(* IEC 61131-3 sources: daoli-st-library/DL_Process (part 16) *)

(* ---- FC_DL_RegisterErrorCalc.st ---- *)
(*
  DL Factory R83 | FC_DL_RegisterErrorCalc
  功能：把纵向与横向套准误差合成偏差幅值与方位角，并按合成允差判定超差。
  开源溯源：无（clean-room 自研，依据公开工艺公式，来源=行业通用公式，许可证=MIT，借鉴点=公式结构）
  规则：R1-R21 全遵守
*)
FUNCTION FC_DL_RegisterErrorCalc : REAL
VAR_INPUT
    fErrMd    : REAL; // 纵向（走料方向）套准误差，正=超前 [mm] / Machine-direction error [mm]
    fErrCd    : REAL; // 横向（幅宽方向）套准误差，正=右偏 [mm] / Cross-direction error [mm]
    fTolMm    : REAL; // 套准允差（合成偏差上限）[mm] / Tolerance on composite error [mm]
    fSpeedMpm : REAL; // 料带走料速度 [m/min] / Web speed [m/min]
END_VAR
VAR_OUTPUT
    fErrComp  : REAL; // 合成偏差幅值 [mm] / Composite error magnitude [mm]
    fErrAngle : REAL; // 误差方位角，0=纵向 90=横向 [°] / Error azimuth [deg]
    xOutTol   : BOOL; // 超差标志（TRUE=超差需调整）/ Out-of-tolerance flag
END_VAR
VAR
    fSq  : REAL; // 误差平方和 [mm²] / Sum of squared errors [mm^2]
    fRad : REAL; // 方位角弧度 [rad] / Azimuth in radians [rad]
    fPi  : REAL := 3.14159265358979; // 圆周率常量，弧度转度用（R19 已引用）/ Pi constant, referenced
END_VAR
// 出口预置：三出口统一预置（R256）
fErrComp := 0.0; fErrAngle := 0.0; xOutTol := FALSE;
// 非有限拦截 + 量纲自检：允差必须为正（R20/R21）
IF NOT (fErrMd > -1.0E30 AND fErrMd < 1.0E30) OR NOT (fErrCd > -1.0E30 AND fErrCd < 1.0E30) OR NOT (fTolMm > -1.0E30 AND fTolMm < 1.0E30) OR NOT (fSpeedMpm > -1.0E30 AND fSpeedMpm < 1.0E30) OR fTolMm <= 0.0 THEN
    FC_DL_RegisterErrorCalc := -1.0; RETURN;   // 哨兵 -1：非有限或允差非正 / Sentinel -1
END_IF
// 合成偏差：欧氏范数，开方前非负闸（R4）
fSq := fErrMd * fErrMd + fErrCd * fErrCd;  // 平方和 [mm²] / Sum of squares [mm^2]
IF fSq >= 0.0 THEN                  // 开方前非负闸 / Gate before square root
    fErrComp := SQRT(fSq);          // 合成偏差 [mm] / Composite error [mm]
ELSE
    fErrComp := 0.0;                // 浮点异常防御缺省 / Float anomaly default
END_IF
// 方位角：纵向分量为分母，显式零闸后取反正切，纯横向走 ±90° 分支
IF ABS(fErrMd) > 1.0E-6 THEN        // 分母零闸（R4/R21）/ Denominator zero gate
    fRad      := ATAN(fErrCd / fErrMd);   // 象限角 [-π/2, π/2] / Quadrant angle [rad]
    fErrAngle := fRad * 180.0 / fPi;      // 转度 [°] / Convert to degrees [deg]
ELSIF fErrCd >= 0.0 THEN
    fErrAngle := 90.0;              // 纯横向正向 [°] / Pure positive cross direction
ELSE
    fErrAngle := -90.0;             // 纯横向负向 [°] / Pure negative cross direction
END_IF
// 超差判定：合成偏差严格大于允差，禁浮点等号比较
xOutTol := fErrComp > fTolMm;       // 超差布尔 / Out-of-tolerance boolean
FC_DL_RegisterErrorCalc := fErrComp; // 返回合成偏差 [mm] / Return composite error [mm]
END_FUNCTION

(* ---- FC_DL_ReOrganicLoadingCalc.st ---- *)
(*
  Component : FC_DL_ReOrganicLoadingCalc
  Category  : DL_Process
  Function  : 有机相稀土负载 g/L = 水相浓度 × 水相流量 / 有机相流量
  Complexity: C2
  开源溯源 : DLF 内部原创（R94 族模板派生）；参考语义来源见 SOURCE_HUNTING_MATRIX.md
  规则遵从 : R1-R16
  契约     : 输入 rAqConcGpl 水相稀土浓度 [g/L]、rFlowAqM3h 水相流量 [m3/h]、rFlowOrgM3h 有机相流量 [m3/h]、
             rLoadMaxGpl 负载上限 [g/L]；输出 rLoadingGpl 有机相负载 [g/L]、rLoadingPct 占上限百分比 [%]、
             xOverLoad 超负载上限（信息级）、xValid 有效标志、nFaultCode 故障码。
  边界     : 有机相流量须 >1.0E-9 [m3/h]（分母下限）；水相浓度须 ≥0；负流量属测量故障判 9801；
             浓度与流量同单位相乘再除，量纲为 g/L，体积流量单位在分子分母相消，无需额外换算系数。
  码位     : 9801 输入非法（故障级）；9802 有机相流量过小（故障级）。
*)
FUNCTION FC_DL_ReOrganicLoadingCalc : BOOL
VAR_INPUT
    rAqConcGpl    : LREAL := 100.0;  // 水相稀土浓度 [g/L] EN: the rare earth concentration of the aqueous phase
    rFlowAqM3h    : LREAL := 5.0;    // 水相体积流量 [m3/h] EN: the volumetric flow of the aqueous phase
    rFlowOrgM3h   : LREAL := 5.0;    // 有机相体积流量 [m3/h] EN: the volumetric flow of the organic phase
    rLoadMaxGpl   : LREAL := 25.0;   // 有机相负载上限 [g/L] EN: the upper limit of the organic phase loading
END_VAR
VAR_OUTPUT
    rLoadingGpl : LREAL;             // 有机相稀土负载 [g/L] EN: the rare earth loading of the organic phase
    rLoadingPct : LREAL;             // 负载占上限的百分比 [%] EN: the loading expressed as a percent of the limit
    xOverLoad   : BOOL;              // 超负载上限（信息级，不置故障） EN: above the loading limit, information class only
    xValid      : BOOL;              // 输出可信标志 EN: the outputs are valid
    nFaultCode  : INT;               // 0=无故障 9801=输入非法 9802=有机相流量过小 EN: zero none, 9801 illegal input, 9802 organic flow too small
END_VAR
VAR
    xFinAll : BOOL;                  // 四输入同时有限 EN: all four inputs are finite
    rDen    : LREAL;                 // 分母（有机相流量） [m3/h] EN: the divisor, the organic phase flow
    rLoad   : LREAL;                 // 负载中间值 [g/L] EN: the interim loading value
END_VAR
VAR CONSTANT
    DL_ROL_Z       : LREAL := 0.0;    // 浮点零常量 EN: the floating point zero constant
    DL_ROL_HUNDRED : LREAL := 100.0;  // 百分数换算系数 EN: the percent conversion factor
    DL_ROL_DEN_MIN : LREAL := 1.0E-9; // 分母绝对值下限 [m3/h] EN: the lower bound of the divisor magnitude
    DL_ROL_C_BAD   : INT := 9801;     // 输入非法 EN: an illegal input
    DL_ROL_C_DEN   : INT := 9802;     // 有机相流量过小 EN: the organic phase flow is too small
END_VAR

// 段1｜出口预置
FC_DL_ReOrganicLoadingCalc := FALSE;   // 返回值预置假 EN: preset the return value to false
rLoadingGpl := DL_ROL_Z;               // 负载预置零 [g/L] EN: preset the loading to zero
rLoadingPct := DL_ROL_Z;               // 负载百分比预置零 [%] EN: preset the loading percent to zero
xOverLoad := FALSE;                    // 超限标志预置假 EN: preset the overload flag to false
xValid := FALSE;                       // 有效标志预置假 EN: preset the validity flag to false
nFaultCode := 0;                       // 故障码预置零 EN: preset the fault code to zero

// 段2｜非有限闸：四个浮点入参全列（上限参与百分比判据，漏则超限判据静默失效）
xFinAll := (rAqConcGpl = rAqConcGpl) AND ((rAqConcGpl - rAqConcGpl) = DL_ROL_Z)
        AND (rFlowAqM3h = rFlowAqM3h) AND ((rFlowAqM3h - rFlowAqM3h) = DL_ROL_Z)
        AND (rFlowOrgM3h = rFlowOrgM3h) AND ((rFlowOrgM3h - rFlowOrgM3h) = DL_ROL_Z)
        AND (rLoadMaxGpl = rLoadMaxGpl) AND ((rLoadMaxGpl - rLoadMaxGpl) = DL_ROL_Z);         // 四输入有限性 EN: the finiteness of all four inputs
IF NOT xFinAll THEN                                                                          // 非有限出口 EN: leave early on a non finite input
    nFaultCode := DL_ROL_C_BAD;                                                              // 输入非法码 EN: the illegal input code
    RETURN;                                                                                  // 早退 EN: return early
END_IF

// 段3｜域闸：浓度非负、两流量非负，有机相流量为分母须过下限
rDen := rFlowOrgM3h;                                                                         // 取分母 [m3/h] EN: take the divisor
IF (rAqConcGpl < DL_ROL_Z) OR (rFlowAqM3h < DL_ROL_Z) OR (ABS(rDen) < DL_ROL_DEN_MIN) THEN   // 域闸 EN: the domain gate
    nFaultCode := DL_ROL_C_DEN;                                                              // 流量或域非法码 EN: the flow or domain code
    RETURN;                                                                                  // 早退 EN: return early
END_IF

// 段4｜主体：负载 = 浓度 × 水相流量 / 有机相流量
rLoad := (rAqConcGpl * rFlowAqM3h) / rDen;                                                   // 负载 [g/L] EN: the organic phase loading
IF (rLoad <> rLoad) OR (rLoad < DL_ROL_Z) THEN                                               // 结果复检：非有限或负 EN: recheck for a non finite or negative result
    nFaultCode := DL_ROL_C_BAD;                                                              // 复检失败码 EN: the recheck failure code
    RETURN;                                                                                  // 早退，出口保持零哨兵 EN: return early with the zero sentinel
END_IF

// 段5｜出口：百分比仅在限值 >0 时计算，否则以 0 表达不可比
rLoadingGpl := rLoad;                                                                        // 负载出口 [g/L] EN: the loading output
IF rLoadMaxGpl > DL_ROL_Z THEN                                                               // 限值有效性 EN: the limit is usable
    rLoadingPct := (rLoad / rLoadMaxGpl) * DL_ROL_HUNDRED;                                   // 占限百分比 [%] EN: the percent of the limit
ELSE
    rLoadingPct := DL_ROL_Z;                                                                 // 限值无效时给零 [%] EN: give zero when the limit is unusable
END_IF
xOverLoad := (rLoadMaxGpl > DL_ROL_Z) AND (rLoad > rLoadMaxGpl);                             // 超限判据（信息级） EN: the overload test, information class only
xValid := TRUE;                                                                              // 结果可信 EN: the results are valid
FC_DL_ReOrganicLoadingCalc := TRUE;                                                          // 返回真 EN: return true
END_FUNCTION

(* ---- FC_DL_RePhaseRatioCalc.st ---- *)
(*
  Component : FC_DL_RePhaseRatioCalc
  Category  : DL_Process
  Function  : 相比 O/A、两相总流量核算与总流量一致性校验
  Complexity: C2
  开源溯源 : DLF 内部原创（R94 族模板派生）；参考语义来源见 SOURCE_HUNTING_MATRIX.md
  规则遵从 : R1-R16
  契约     : 输入 rFlowOrgM3h 有机相流量 [m3/h]、rFlowAqM3h 水相流量 [m3/h]、
             rFlowTotalMeasM3h 实测混合前总流量 [m3/h]、rTotalTolPct 总流量相对容差 [%]；
             输出 rRatioOA 相比 [-]、rFlowTotalM3h 计算总流量 [m3/h]、rDevPct 相对偏差 [%]、
             xTotalMatch 总流量一致、xValid 有效标志、nFaultCode 故障码。
  边界     : 水相流量为分母须 >1.0E-9 [m3/h]；两流量均须 ≥0；总流量容差须在 (0, 100] [%] 内，
             否则判 9803（容差非法会使一致性判据恒真或恒假，属组态域闸缺失）；
             相对偏差以计算总流量为分母，故须先证计算总流量 >1.0E-9。
  码位     : 9801 输入非法（故障级）；9802 水相流量过小（故障级）；9803 容差越域（故障级）。
*)
FUNCTION FC_DL_RePhaseRatioCalc : BOOL
VAR_INPUT
    rFlowOrgM3h       : LREAL := 5.0;    // 有机相体积流量 [m3/h] EN: the volumetric flow of the organic phase
    rFlowAqM3h        : LREAL := 5.0;    // 水相体积流量 [m3/h] EN: the volumetric flow of the aqueous phase
    rFlowTotalMeasM3h : LREAL := 10.0;   // 实测总流量（混合前两路之和） [m3/h] EN: the measured total flow of both phases before mixing
    rTotalTolPct      : LREAL := 2.0;    // 总流量相对容差 [%] EN: the relative tolerance of the total flow
END_VAR
VAR_OUTPUT
    rRatioOA     : LREAL;                // 相比 O/A [-] EN: the organic to aqueous phase ratio
    rFlowTotalM3h: LREAL;                // 计算总流量 [m3/h] EN: the computed total flow
    rDevPct      : LREAL;                // 实测相对计算值的偏差 [%] EN: the deviation of the measurement from the computed total
    xTotalMatch  : BOOL;                 // 总流量一致（在容差内） EN: the total flow agrees within the tolerance
    xValid       : BOOL;                 // 输出可信标志 EN: the outputs are valid
    nFaultCode   : INT;                  // 0=无故障 9801=输入非法 9802=水相流量过小 9803=容差越域 EN: zero none, 9801 illegal input, 9802 aqueous flow too small, 9803 tolerance out of range
END_VAR
VAR
    xFinAll   : BOOL;                    // 四输入同时有限 EN: all four inputs are finite
    xNegFlow  : BOOL;                    // 存在负流量 EN: some flow is negative
    rDen      : LREAL;                   // 分母（水相流量） [m3/h] EN: the divisor, the aqueous phase flow
    rTotal    : LREAL;                   // 计算总流量中间值 [m3/h] EN: the interim computed total flow
    rDev      : LREAL;                   // 偏差中间值 [%] EN: the interim deviation value
END_VAR
VAR CONSTANT
    DL_RPR_Z       : LREAL := 0.0;       // 浮点零常量 EN: the floating point zero constant
    DL_RPR_HUNDRED : LREAL := 100.0;     // 百分数换算系数 EN: the percent conversion factor
    DL_RPR_DEN_MIN : LREAL := 1.0E-9;    // 分母绝对值下限 [m3/h] EN: the lower bound of the divisor magnitude
    DL_RPR_C_BAD   : INT := 9801;        // 输入非法 EN: an illegal input
    DL_RPR_C_DEN   : INT := 9802;        // 水相流量过小 EN: the aqueous phase flow is too small
    DL_RPR_C_TOL   : INT := 9803;        // 容差越域 EN: the tolerance is out of range
END_VAR

// 段1｜出口预置
FC_DL_RePhaseRatioCalc := FALSE;   // 返回值预置假 EN: preset the return value to false
rRatioOA := DL_RPR_Z;              // 相比预置零 [-] EN: preset the phase ratio to zero
rFlowTotalM3h := DL_RPR_Z;         // 总流量预置零 [m3/h] EN: preset the total flow to zero
rDevPct := DL_RPR_Z;               // 偏差预置零 [%] EN: preset the deviation to zero
xTotalMatch := FALSE;              // 一致标志预置假 EN: preset the agreement flag to false
xValid := FALSE;                   // 有效标志预置假 EN: preset the validity flag to false
nFaultCode := 0;                   // 故障码预置零 EN: preset the fault code to zero

// 段2｜非有限闸：四个浮点入参全列，容差虽为限值但不入闸则一致性判据可被 NaN 击穿
xFinAll := (rFlowOrgM3h = rFlowOrgM3h) AND ((rFlowOrgM3h - rFlowOrgM3h) = DL_RPR_Z)
        AND (rFlowAqM3h = rFlowAqM3h) AND ((rFlowAqM3h - rFlowAqM3h) = DL_RPR_Z)
        AND (rFlowTotalMeasM3h = rFlowTotalMeasM3h) AND ((rFlowTotalMeasM3h - rFlowTotalMeasM3h) = DL_RPR_Z)
        AND (rTotalTolPct = rTotalTolPct) AND ((rTotalTolPct - rTotalTolPct) = DL_RPR_Z);   // 四输入有限性 EN: the finiteness of all four inputs
IF NOT xFinAll THEN                                                                          // 非有限出口 EN: leave early on a non finite input
    nFaultCode := DL_RPR_C_BAD;                                                              // 输入非法码 EN: the illegal input code
    RETURN;                                                                                  // 早退 EN: return early
END_IF

// 段3｜域闸：两流量非负、水相流量过分母下限、容差落在 (0,100] 域内
xNegFlow := (rFlowOrgM3h < DL_RPR_Z) OR (rFlowAqM3h < DL_RPR_Z);                             // 负流量判据 EN: the negative flow test
rDen := rFlowAqM3h;                                                                          // 取分母 [m3/h] EN: take the divisor
IF xNegFlow OR (ABS(rDen) < DL_RPR_DEN_MIN) THEN                                             // 流量域闸 EN: the flow domain gate
    nFaultCode := DL_RPR_C_DEN;                                                              // 流量非法码 EN: the flow code
    RETURN;                                                                                  // 早退 EN: return early
END_IF
IF (rTotalTolPct <= DL_RPR_Z) OR (rTotalTolPct > DL_RPR_HUNDRED) THEN                        // 容差域闸 EN: the tolerance domain gate
    nFaultCode := DL_RPR_C_TOL;                                                              // 容差越域码 EN: the tolerance code
    RETURN;                                                                                  // 早退 EN: return early
END_IF

// 段4｜主体：相比与计算总流量
rTotal := rFlowOrgM3h + rFlowAqM3h;                                                          // 计算总流量 [m3/h] EN: the computed total flow
rRatioOA := rFlowOrgM3h / rDen;                                                              // 相比 O/A [-] EN: the phase ratio
rFlowTotalM3h := rTotal;                                                                     // 总流量出口 [m3/h] EN: the total flow output

// 段5｜一致性校验：偏差以计算总流量为分母，先证其过下限
IF ABS(rTotal) < DL_RPR_DEN_MIN THEN                                                         // 总流量分母下限 EN: the total flow divisor gate
    rDev := DL_RPR_Z;                                                                        // 偏差给零 [%] EN: give a zero deviation
    xTotalMatch := FALSE;                                                                    // 不可比，判不一致 EN: not comparable, report a mismatch
ELSE
    rDev := (rFlowTotalMeasM3h - rTotal) / rTotal * DL_RPR_HUNDRED;                         // 相对偏差 [%] EN: the relative deviation
    xTotalMatch := ABS(rDev) <= rTotalTolPct;                                                // 容差比较 EN: the tolerance comparison
END_IF
rDevPct := rDev;                                                                             // 偏差出口 [%] EN: the deviation output
xValid := TRUE;                                                                              // 结果可信 EN: the results are valid
FC_DL_RePhaseRatioCalc := TRUE;                                                              // 返回真 EN: return true
END_FUNCTION

(* ---- FC_DL_ReProductPurityCalc.st ---- *)
(*
  Component : FC_DL_ReProductPurityCalc
  Category  : DL_Process
  Function  : 产品纯度 = (1 - Σ杂质/总量) × 100，并给出合格判定
  Complexity: C2
  开源溯源 : DLF 内部原创（R94 族模板派生）；参考语义来源见 SOURCE_HUNTING_MATRIX.md
  规则遵从 : R1-R16
  契约     : 输入 afImpPpm 杂质浓度定长数组 [ppm]（ARRAY[0..7]，R15 显式定长）、nImpCount 有效杂质个数 [个]、
             rTotalPpm 总量基准 [ppm]、rPuritySpecPct 纯度合格下限 [%]；
             输出 rImpSumPpm 杂质合计 [ppm]、rPurityPct 产品纯度 [%]、xPass 合格、
             xClamped 本拍钳位、xValid 有效标志、nFaultCode 故障码。
  边界     : 数组固定 8 元素，nImpCount 须在 0..8 内，越界判 9803 并拒绝访问；总量基准须 >1.0E-9 [ppm] 判 9802；
             任一有效元素非有限判 9801；纯度钳位 0~100 [%]；杂质合计超过总量时纯度钳到零并置 xClamped。
  码位     : 9801 元素非有限（故障级）；9802 总量基准过小（故障级）；9803 杂质个数越界（故障级）。
*)
FUNCTION FC_DL_ReProductPurityCalc : BOOL
VAR_INPUT
    afImpPpm      : ARRAY[0..7] OF LREAL;   // 杂质浓度定长数组，未用槽填零 [ppm] EN: the fixed impurity concentration array, unused slots hold zero
    nImpCount     : INT := 8;               // 有效杂质元素个数 [个] EN: the number of valid impurity elements
    rTotalPpm     : LREAL := 1000000.0;     // 总量基准（纯度分母） [ppm] EN: the total amount used as the purity divisor
    rPuritySpecPct: LREAL := 99.5;          // 纯度合格下限 [%] EN: the lower acceptance limit of the product purity
END_VAR
VAR_OUTPUT
    rImpSumPpm : LREAL;                     // 有效杂质合计 [ppm] EN: the sum of the valid impurities
    rPurityPct : LREAL;                     // 产品纯度，域 0~100 [%] EN: the product purity clamped to zero through one hundred
    xPass      : BOOL;                      // 纯度合格判定 EN: the purity acceptance verdict
    xClamped   : BOOL;                      // 本拍发生钳位 EN: a clamp occurred in this cycle
    xValid     : BOOL;                      // 输出可信标志 EN: the outputs are valid
    nFaultCode : INT;                       // 0=无故障 9801=元素非有限 9802=总量过小 9803=个数越界 EN: zero none, 9801 non finite element, 9802 total too small, 9803 count out of range
END_VAR
VAR
    xFinAll  : BOOL;                        // 全部元素有限（仅扫有效区） EN: every scanned element is finite
    xFinEl   : BOOL;                        // 单元素有限性 EN: the finiteness of one element
    i        : INT;                         // 杂质数组循环索引 [个] EN: the impurity array loop index
    nScan    : INT;                         // 实际扫描个数 [个] EN: the effective scan count
    rSum     : LREAL;                       // 杂质累加器 [ppm] EN: the impurity accumulator
    rRatio   : LREAL;                       // 杂质占总量比例 [-] EN: the impurity fraction of the total
    rPur     : LREAL;                       // 纯度中间值 [%] EN: the interim purity value
END_VAR
VAR CONSTANT
    DL_RPP_Z        : LREAL := 0.0;         // 浮点零常量 EN: the floating point zero constant
    DL_RPP_ONE      : LREAL := 1.0;         // 浮点壹常量 EN: the floating point one constant
    DL_RPP_HUNDRED  : LREAL := 100.0;       // 百分数换算系数 EN: the percent conversion factor
    DL_RPP_IDX_MAX  : INT := 7;             // 数组上界索引 [个] EN: the array upper bound index
    DL_RPP_CNT_MAX  : INT := 8;             // 允许的杂质个数上限 [个] EN: the allowed upper bound of the impurity count
    DL_RPP_C_BAD    : INT := 9801;          // 元素非有限 EN: a non finite element
    DL_RPP_C_TOTAL  : INT := 9802;          // 总量过小 EN: the total amount is too small
    DL_RPP_C_INDEX  : INT := 9803;          // 杂质个数越界 EN: the impurity count is out of range
END_VAR

// 段1｜出口预置
FC_DL_ReProductPurityCalc := FALSE;   // 返回值预置假 EN: preset the return value to false
rImpSumPpm := DL_RPP_Z;               // 杂质合计预置零 [ppm] EN: preset the impurity sum to zero
rPurityPct := DL_RPP_Z;               // 纯度预置零 [%] EN: preset the purity to zero
xPass := FALSE;                       // 合格标志预置假 EN: preset the acceptance flag to false
xClamped := FALSE;                    // 钳位标志预置假 EN: preset the clamp flag to false
xValid := FALSE;                      // 有效标志预置假 EN: preset the validity flag to false
nFaultCode := 0;                      // 故障码预置零 EN: preset the fault code to zero

// 段2｜非有限闸：三个标量入参全列（合格下限参与出口判据）
xFinAll := (rTotalPpm = rTotalPpm) AND ((rTotalPpm - rTotalPpm) = DL_RPP_Z)
        AND (rPuritySpecPct = rPuritySpecPct) AND ((rPuritySpecPct - rPuritySpecPct) = DL_RPP_Z);   // 标量有限性 EN: the finiteness of the scalar inputs
IF NOT xFinAll THEN                                                                                 // 非有限出口 EN: leave early on a non finite input
    nFaultCode := DL_RPP_C_BAD;                                                                     // 输入非法码 EN: the illegal input code
    RETURN;                                                                                         // 早退 EN: return early
END_IF

// 段3｜域闸：杂质个数在 0..8 内（越界一律拒绝访问，不做截断放行）
IF (nImpCount < 0) OR (nImpCount > DL_RPP_CNT_MAX) OR (ABS(rTotalPpm) < 1.0E-9) THEN                  // 索引与分母域闸 EN: the index and divisor domain gate
    IF (nImpCount < 0) OR (nImpCount > DL_RPP_CNT_MAX) THEN                                          // 区分越界与分母两类成因 EN: separate the index cause from the divisor cause
        nFaultCode := DL_RPP_C_INDEX;                                                                // 个数越界码 EN: the count out of range code
    ELSE
        nFaultCode := DL_RPP_C_TOTAL;                                                                // 总量过小码 EN: the total too small code
    END_IF
    RETURN;                                                                                          // 早退 EN: return early
END_IF

// 段4｜主体：扫有效区累加杂质，逐元素过非有限闸（非有限拒收，不参与累加）
rSum := DL_RPP_Z;                                                                                    // 累加器清零 [ppm] EN: clear the accumulator
nScan := nImpCount;                                                                                  // 扫描个数 [个] EN: the scan count
xFinAll := TRUE;                                                                                     // 假定全部有限 EN: assume every element is finite
FOR i := 0 TO nScan - 1 DO                                                                           // 定长数组循环，nScan 已证 ≤8 EN: the fixed array loop, the count is proven at most eight
    IF (i >= 0) AND (i <= DL_RPP_IDX_MAX) THEN                                                       // 逐元素双边界校验 EN: the per element bound check
        xFinEl := (afImpPpm[i] = afImpPpm[i]) AND ((afImpPpm[i] - afImpPpm[i]) = DL_RPP_Z);          // 元素有限性 EN: the element finiteness
        IF xFinEl THEN                                                                               // 有限才累加 EN: accumulate only finite values
            rSum := rSum + afImpPpm[i];                                                              // 累加杂质 [ppm] EN: accumulate the impurity
        ELSE
            xFinAll := FALSE;                                                                        // 记非有限 EN: mark the non finite element
        END_IF
    END_IF
END_FOR
IF NOT xFinAll THEN                                                                                  // 存在非有限元素 EN: some element is not finite
    nFaultCode := DL_RPP_C_BAD;                                                                      // 元素非有限码 EN: the non finite element code
    rImpSumPpm := DL_RPP_Z;                                                                          // 合计复位零哨兵 [ppm] EN: reset the sum to the zero sentinel
    RETURN;                                                                                          // 早退 EN: return early
END_IF

// 段5｜纯度：先算比例再钳位（负比例来自负杂质输入，属组态错误，钳零并留痕）
rRatio := rSum / rTotalPpm;                                                                          // 杂质比例，分母已过下限 [-] EN: the impurity fraction, the divisor passed the gate
rPur := (DL_RPP_ONE - rRatio) * DL_RPP_HUNDRED;                                                      // 纯度 [%] EN: the purity
IF rPur < DL_RPP_Z THEN                                                                              // 下钳位 EN: clamp the lower bound
    rPur := DL_RPP_Z;                                                                                // 钳到零 [%] EN: clamp to zero
    xClamped := TRUE;                                                                                // 置钳位标志 EN: raise the clamp flag
END_IF
IF rPur > DL_RPP_HUNDRED THEN                                                                        // 上钳位 EN: clamp the upper bound
    rPur := DL_RPP_HUNDRED;                                                                          // 钳到一百 [%] EN: clamp to one hundred
    xClamped := TRUE;                                                                                // 置钳位标志 EN: raise the clamp flag
END_IF

// 段6｜出口：名实双出口同源，合格判定用钳位后的纯度
rImpSumPpm := rSum;                                                                                  // 合计出口 [ppm] EN: the impurity sum output
rPurityPct := rPur;                                                                                  // 纯度出口 [%] EN: the purity output
xPass := rPur >= rPuritySpecPct;                                                                     // 合格判定 EN: the acceptance verdict
xValid := TRUE;                                                                                      // 结果可信 EN: the results are valid
FC_DL_ReProductPurityCalc := TRUE;                                                                   // 返回真 EN: return true
END_FUNCTION

(* ---- FC_DL_ReSaponificationRateCalc.st ---- *)
(*
  Component : FC_DL_ReSaponificationRateCalc
  Category  : DL_Process
  Function  : 皂化率 = 实际皂化碱量 / 理论碱量 × 100，并钳位到 0~100
  Complexity: C2
  开源溯源 : DLF 内部原创（R94 族模板派生）；参考语义来源见 SOURCE_HUNTING_MATRIX.md
  规则遵从 : R1-R16
  契约     : 输入 rAlkaliActual 实际皂化碱量 [kg/h]、rAlkaliTheory 理论皂化碱量 [kg/h]、
             rRateHighLimit 判定上限 [%]；输出 rRateRaw 未钳位皂化率 [%]、rRatePct 钳位后皂化率 [%]、
             xClamped 钳位发生标志、xOverRate 超判定上限标志、xValid 有效标志、nFaultCode 故障码。
  边界     : 理论碱量须 >1.0E-9 [kg/h]，否则判 9802；实际碱量为负判 9801（负投加不可能，属测量故障）；
             钳位范围 0~100 [%] 为物理可实现域；xClamped 只表达本拍是否发生钳位，不置故障。
  码位     : 9801 输入非法（故障级）；9802 理论碱量过小（故障级）。信息级钳位不派码，由 xClamped 表达。
*)
FUNCTION FC_DL_ReSaponificationRateCalc : BOOL
VAR_INPUT
    rAlkaliActual   : LREAL := 10.0;   // 实际皂化碱量 [kg/h] EN: the actual alkali mass flow used for saponification
    rAlkaliTheory   : LREAL := 12.0;   // 理论皂化碱量 [kg/h] EN: the theoretical alkali mass flow required by stoichiometry
    rRateHighLimit  : LREAL := 100.0;  // 皂化率合格上限 [%] EN: the upper limit of an acceptable saponification rate
END_VAR
VAR_OUTPUT
    rRateRaw   : LREAL;                // 未钳位皂化率 [%] EN: the saponification rate before clamping
    rRatePct   : LREAL;                // 钳位后皂化率，域 0~100 [%] EN: the saponification rate clamped to zero through one hundred
    xClamped   : BOOL;                 // 本拍发生钳位 EN: a clamp occurred in this cycle
    xOverRate  : BOOL;                 // 超判定上限（信息级） EN: the rate exceeds the upper limit, an information class flag
    xValid     : BOOL;                 // 输出可信标志 EN: the outputs are valid
    nFaultCode : INT;                  // 0=无故障 9801=输入非法 9802=理论碱量过小 EN: zero none, 9801 illegal input, 9802 theoretical alkali too small
END_VAR
VAR
    xFinAll  : BOOL;                   // 三输入同时有限 EN: all three inputs are finite
    xNegAct  : BOOL;                   // 实际碱量为负 EN: the actual alkali flow is negative
    rDen     : LREAL;                  // 分母（理论碱量） [kg/h] EN: the divisor, the theoretical alkali flow
    rRaw     : LREAL;                  // 皂化率中间值 [%] EN: the interim saponification rate
    rClamp   : LREAL;                  // 钳位结果 [%] EN: the clamped result
END_VAR
VAR CONSTANT
    DL_SSR_Z       : LREAL := 0.0;     // 浮点零常量 EN: the floating point zero constant
    DL_SSR_HUNDRED : LREAL := 100.0;   // 百分数换算系数 EN: the percent conversion factor
    DL_SSR_DEN_MIN : LREAL := 1.0E-9;  // 分母绝对值下限 [kg/h] EN: the lower bound of the divisor magnitude
    DL_SSR_C_BAD   : INT := 9801;      // 输入非法 EN: an illegal input
    DL_SSR_C_DEN   : INT := 9802;      // 理论碱量过小 EN: the theoretical alkali flow is too small
END_VAR

// 段1｜出口预置
FC_DL_ReSaponificationRateCalc := FALSE;   // 返回值预置假 EN: preset the return value to false
rRateRaw := DL_SSR_Z;                      // 未钳位皂化率预置零 [%] EN: preset the raw rate to zero
rRatePct := DL_SSR_Z;                      // 钳位皂化率预置零 [%] EN: preset the clamped rate to zero
xClamped := FALSE;                         // 钳位标志预置假 EN: preset the clamp flag to false
xOverRate := FALSE;                        // 超限标志预置假 EN: preset the over rate flag to false
xValid := FALSE;                           // 有效标志预置假 EN: preset the validity flag to false
nFaultCode := 0;                           // 故障码预置零 EN: preset the fault code to zero

// 段2｜非有限闸：三个浮点入参逐一列入（上限限值同样参与判据换算，不可漏）
xFinAll := (rAlkaliActual = rAlkaliActual) AND ((rAlkaliActual - rAlkaliActual) = DL_SSR_Z)
        AND (rAlkaliTheory = rAlkaliTheory) AND ((rAlkaliTheory - rAlkaliTheory) = DL_SSR_Z)
        AND (rRateHighLimit = rRateHighLimit) AND ((rRateHighLimit - rRateHighLimit) = DL_SSR_Z);   // 三输入有限性 EN: the finiteness of all three inputs
IF NOT xFinAll THEN                                                                                  // 非有限出口 EN: leave early on a non finite input
    nFaultCode := DL_SSR_C_BAD;                                                                      // 输入非法码 EN: the illegal input code
    RETURN;                                                                                          // 早退 EN: return early
END_IF

// 段3｜域闸：理论碱量为分母须足够大；实际碱量不得为负（负投加属测量方向故障）
rDen := rAlkaliTheory;                                                                               // 取分母 [kg/h] EN: take the divisor
xNegAct := rAlkaliActual < DL_SSR_Z;                                                                 // 负投加判据 EN: the negative dosing test
IF (ABS(rDen) < DL_SSR_DEN_MIN) OR xNegAct OR (rRateHighLimit <= DL_SSR_Z) THEN                     // 域闸 EN: the domain gate
    nFaultCode := DL_SSR_C_DEN;                                                                      // 分母或域非法码 EN: the divisor or domain code
    RETURN;                                                                                          // 早退 EN: return early
END_IF

// 段4｜主体：raw = 实际 / 理论 × 100，钳位 0~100
rRaw := (rAlkaliActual / rDen) * DL_SSR_HUNDRED;                                                     // 未钳位皂化率 [%] EN: the saponification rate before clamping
rClamp := rRaw;                                                                                      // 钳位工作副本 [%] EN: the working copy for clamping
IF rClamp < DL_SSR_Z THEN                                                                            // 下钳位 EN: clamp the lower bound
    rClamp := DL_SSR_Z;                                                                              // 钳到零 [%] EN: clamp to zero
    xClamped := TRUE;                                                                                // 置钳位标志 EN: raise the clamp flag
END_IF
IF rClamp > DL_SSR_HUNDRED THEN                                                                      // 上钳位 EN: clamp the upper bound
    rClamp := DL_SSR_HUNDRED;                                                                        // 钳到一百 [%] EN: clamp to one hundred
    xClamped := TRUE;                                                                                // 置钳位标志 EN: raise the clamp flag
END_IF

// 段5｜出口：名实双出口同源赋值，超限为信息级不置故障
rRateRaw := rRaw;                                                                                    // 未钳位出口 [%] EN: the raw rate output
rRatePct := rClamp;                                                                                  // 钳位出口 [%] EN: the clamped rate output
xOverRate := rClamp > rRateHighLimit;                                                                // 超判定上限（信息级） EN: above the acceptance limit, information class only
xValid := TRUE;                                                                                      // 结果可信 EN: the results are valid
FC_DL_ReSaponificationRateCalc := TRUE;                                                              // 返回真 EN: return true
END_FUNCTION

(* ---- FC_DL_ReStageEfficiencyCalc.st ---- *)
(*
  Component : FC_DL_ReStageEfficiencyCalc
  Category  : DL_Process
  Function  : 单级萃取效率 = 实际萃取量 / 平衡萃取量 × 100，并钳位到 0~100
  Complexity: C2
  开源溯源 : DLF 内部原创（R94 族模板派生）；参考语义来源见 SOURCE_HUNTING_MATRIX.md
  规则遵从 : R1-R16
  契约     : 输入 rActualExtractGpl 实际萃取量 [g/L]、rEquilExtractGpl 平衡萃取量 [g/L]、
             rEffHighPct 效率合格下限 [%]；输出 rEffRawPct 未钳位效率 [%]、rEffPct 钳位后效率 [%]、
             xClamped 本拍钳位、xEffLow 效率低于合格下限（信息级）、xValid 有效标志、nFaultCode 故障码。
  边界     : 平衡萃取量为分母须 >1.0E-9 [g/L]；实际萃取量为负判 9801（负萃取属测量方向故障）；
             钳位域 0~100 [%]；xEffLow 为信息级，不置故障，仅当效率低于合格下限时置位。
  码位     : 9801 输入非法（故障级）；9802 平衡萃取量过小（故障级）。
*)
FUNCTION FC_DL_ReStageEfficiencyCalc : BOOL
VAR_INPUT
    rActualExtractGpl : LREAL := 8.0;    // 单级实际萃取量 [g/L] EN: the rare earth mass actually extracted in one stage
    rEquilExtractGpl  : LREAL := 10.0;   // 单级平衡萃取量 [g/L] EN: the rare earth mass extracted at equilibrium in one stage
    rEffHighPct       : LREAL := 90.0;   // 单级效率合格下限 [%] EN: the lower acceptance limit of the single stage efficiency
END_VAR
VAR_OUTPUT
    rEffRawPct : LREAL;                  // 未钳位单级效率 [%] EN: the single stage efficiency before clamping
    rEffPct    : LREAL;                  // 钳位后单级效率，域 0~100 [%] EN: the single stage efficiency clamped to zero through one hundred
    xClamped   : BOOL;                   // 本拍发生钳位 EN: a clamp occurred in this cycle
    xEffLow    : BOOL;                   // 效率低于合格下限（信息级） EN: the efficiency is below the acceptance limit, information class only
    xValid     : BOOL;                   // 输出可信标志 EN: the outputs are valid
    nFaultCode : INT;                    // 0=无故障 9801=输入非法 9802=平衡量过小 EN: zero none, 9801 illegal input, 9802 equilibrium mass too small
END_VAR
VAR
    xFinAll : BOOL;                      // 三输入同时有限 EN: all three inputs are finite
    rDen    : LREAL;                     // 分母（平衡萃取量） [g/L] EN: the divisor, the equilibrium extracted mass
    rRaw    : LREAL;                     // 效率中间值 [%] EN: the interim efficiency value
    rClamp  : LREAL;                     // 钳位工作副本 [%] EN: the working copy for clamping
END_VAR
VAR CONSTANT
    DL_RSE_Z       : LREAL := 0.0;       // 浮点零常量 EN: the floating point zero constant
    DL_RSE_HUNDRED : LREAL := 100.0;     // 百分数换算系数 EN: the percent conversion factor
    DL_RSE_DEN_MIN : LREAL := 1.0E-9;    // 分母绝对值下限 [g/L] EN: the lower bound of the divisor magnitude
    DL_RSE_C_BAD   : INT := 9801;        // 输入非法 EN: an illegal input
    DL_RSE_C_DEN   : INT := 9802;        // 平衡萃取量过小 EN: the equilibrium mass is too small
END_VAR

// 段1｜出口预置
FC_DL_ReStageEfficiencyCalc := FALSE;   // 返回值预置假 EN: preset the return value to false
rEffRawPct := DL_RSE_Z;                 // 未钳位效率预置零 [%] EN: preset the raw efficiency to zero
rEffPct := DL_RSE_Z;                    // 钳位效率预置零 [%] EN: preset the clamped efficiency to zero
xClamped := FALSE;                      // 钳位标志预置假 EN: preset the clamp flag to false
xEffLow := FALSE;                       // 低效标志预置假 EN: preset the low efficiency flag to false
xValid := FALSE;                        // 有效标志预置假 EN: preset the validity flag to false
nFaultCode := 0;                        // 故障码预置零 EN: preset the fault code to zero

// 段2｜非有限闸：三输入全列（合格下限参与出口判据，漏则低效判据失效）
xFinAll := (rActualExtractGpl = rActualExtractGpl) AND ((rActualExtractGpl - rActualExtractGpl) = DL_RSE_Z)
        AND (rEquilExtractGpl = rEquilExtractGpl) AND ((rEquilExtractGpl - rEquilExtractGpl) = DL_RSE_Z)
        AND (rEffHighPct = rEffHighPct) AND ((rEffHighPct - rEffHighPct) = DL_RSE_Z);   // 三输入有限性 EN: the finiteness of all three inputs
IF NOT xFinAll THEN                                                                     // 非有限出口 EN: leave early on a non finite input
    nFaultCode := DL_RSE_C_BAD;                                                         // 输入非法码 EN: the illegal input code
    RETURN;                                                                             // 早退 EN: return early
END_IF

// 段3｜域闸：实际量非负、平衡量过分母下限
rDen := rEquilExtractGpl;                                                               // 取分母 [g/L] EN: take the divisor
IF (rActualExtractGpl < DL_RSE_Z) OR (ABS(rDen) < DL_RSE_DEN_MIN) THEN                  // 域闸 EN: the domain gate
    nFaultCode := DL_RSE_C_DEN;                                                         // 分母或域非法码 EN: the divisor or domain code
    RETURN;                                                                             // 早退 EN: return early
END_IF

// 段4｜主体：eff = 实际 / 平衡 × 100
rRaw := (rActualExtractGpl / rDen) * DL_RSE_HUNDRED;                                    // 未钳位效率 [%] EN: the efficiency before clamping
rClamp := rRaw;                                                                         // 钳位工作副本 [%] EN: the working copy for clamping
IF rClamp < DL_RSE_Z THEN                                                               // 下钳位 EN: clamp the lower bound
    rClamp := DL_RSE_Z;                                                                 // 钳到零 [%] EN: clamp to zero
    xClamped := TRUE;                                                                   // 置钳位标志 EN: raise the clamp flag
END_IF
IF rClamp > DL_RSE_HUNDRED THEN                                                         // 上钳位 EN: clamp the upper bound
    rClamp := DL_RSE_HUNDRED;                                                           // 钳到一百 [%] EN: clamp to one hundred
    xClamped := TRUE;                                                                   // 置钳位标志 EN: raise the clamp flag
END_IF

// 段5｜出口：名实双出口同源赋值；低效为信息级，不置故障
rEffRawPct := rRaw;                                                                     // 未钳位出口 [%] EN: the raw efficiency output
rEffPct := rClamp;                                                                      // 钳位出口 [%] EN: the clamped efficiency output
xEffLow := rClamp < rEffHighPct;                                                        // 低效判据（信息级） EN: the low efficiency test, information class only
xValid := TRUE;                                                                         // 结果可信 EN: the results are valid
FC_DL_ReStageEfficiencyCalc := TRUE;                                                    // 返回真 EN: return true
END_FUNCTION

(* ---- FC_DL_ReStripAcidDosageCalc.st ---- *)
(*
  Component : FC_DL_ReStripAcidDosageCalc
  Category  : DL_Process
  Function  : 反萃酸耗核算：稀土摩尔量 × 当量系数 → 纯酸 kg/h 与所需酸液体积流量、酸浓度校核
  Complexity: C2
  开源溯源 : DLF 内部原创（R94 族模板派生）；参考语义来源见 SOURCE_HUNTING_MATRIX.md
  规则遵从 : R1-R16
  契化     : 输入 rOrgReConcGpl 负载有机相稀土浓度 [g/L]、rFlowOrgM3h 有机相流量 [m3/h]、
             rReMolWeight 稀土平均摩尔质量 [g/mol]、rAcidEquiv 每摩尔稀土耗酸当量 [mol/mol]、
             rAcidMolWeight 酸摩尔质量 [g/mol]、rAcidConcGpl 配酸浓度 [g/L]；
             输出 rReMolH 稀土摩尔流率 [mol/h]、rAcidKgH 纯酸耗量 [kg/h]、rAcidSolM3h 所需酸液体积流量 [m3/h]、
             rAcidExcessPct 实际配酸相对需求的富余率 [%]、xConcOk 浓度配置可行、xValid 有效标志、nFaultCode 故障码。
  边界     : 单位链：g/L × m3/h = 1000 g/h，再除 g/mol 得 mol/h，故 mol/h = 浓度 × 流量 × 1000 / 摩尔质量；
             纯酸 kg/h = mol/h × 当量 × (g/mol) / 1000；g/L 与 kg/m3 数值相等，故酸液 m3/h = kg/h ÷ (g/L)；
             所有摩尔质量与当量须 >1.0E-6，配酸浓度须 >1.0E-9 [g/L]，否则判 9802；
             xConcOk 的判据是「配酸浓度足以在有机相流量同等体积下供足酸量」，不足为信息级告警。
  码位     : 9801 输入非法（故障级）；9802 摩尔质量/当量/配酸浓度越域（故障级）。
*)
FUNCTION FC_DL_ReStripAcidDosageCalc : BOOL
VAR_INPUT
    rOrgReConcGpl   : LREAL := 20.0;    // 负载有机相稀土浓度 [g/L] EN: the rare earth concentration of the loaded organic phase
    rFlowOrgM3h     : LREAL := 5.0;     // 有机相体积流量 [m3/h] EN: the volumetric flow of the organic phase
    rReMolWeight    : LREAL := 140.0;   // 稀土元素平均摩尔质量 [g/mol] EN: the average molar mass of the rare earth element
    rAcidEquiv      : LREAL := 3.0;     // 每摩尔稀土耗酸当量 [mol/mol] EN: the acid equivalents consumed per mole of rare earth
    rAcidMolWeight  : LREAL := 36.46;   // 酸摩尔质量（盐酸缺省） [g/mol] EN: the molar mass of the acid, hydrochloric by default
    rAcidConcGpl    : LREAL := 200.0;   // 配酸浓度 [g/L] EN: the concentration of the prepared acid solution
END_VAR
VAR_OUTPUT
    rReMolH        : LREAL;             // 稀土摩尔流率 [mol/h] EN: the molar flow of the rare earth
    rAcidKgH       : LREAL;             // 纯酸耗量 [kg/h] EN: the pure acid mass flow required
    rAcidSolM3h    : LREAL;             // 所需酸液体积流量 [m3/h] EN: the acid solution volumetric flow required
    rAcidExcessPct : LREAL;             // 配酸富余率（相对同体积供酸能力） [%] EN: the surplus of the prepared acid against the demand at the same volume
    xConcOk        : BOOL;              // 配酸浓度足以供酸（信息级） EN: the acid concentration is sufficient, information class only
    xValid         : BOOL;              // 输出可信标志 EN: the outputs are valid
    nFaultCode     : INT;               // 0=无故障 9801=输入非法 9802=摩尔质量或浓度越域 EN: zero none, 9801 illegal input, 9802 molar mass or concentration out of range
END_VAR
VAR
    xFinAll  : BOOL;                    // 六输入同时有限 EN: all six inputs are finite
    rMolH    : LREAL;                   // 摩尔流率中间值 [mol/h] EN: the interim molar flow
    rAcidKg  : LREAL;                   // 纯酸流量中间值 [kg/h] EN: the interim pure acid mass flow
    rSolM3h  : LREAL;                   // 酸液流量中间值 [m3/h] EN: the interim acid solution flow
    rSupply  : LREAL;                   // 同等体积下的供酸能力 [kg/h] EN: the acid supply capability at the same volumetric flow
END_VAR
VAR CONSTANT
    DL_RSD_Z      : LREAL := 0.0;       // 浮点零常量 EN: the floating point zero constant
    DL_RSD_K1000  : LREAL := 1000.0;    // 升-立方米与克-千克换算系数 EN: the litre to cubic metre and gram to kilogram factor
    DL_RSD_HUND   : LREAL := 100.0;     // 百分数换算系数 EN: the percent conversion factor
    DL_RSD_MIN    : LREAL := 1.0E-6;    // 摩尔质量与当量的下限 EN: the lower bound of the molar mass and equivalents
    DL_RSD_C_BAD  : INT := 9801;        // 输入非法 EN: an illegal input
    DL_RSD_C_RANGE: INT := 9802;        // 摩尔质量或配酸浓度越域 EN: the molar mass or the acid concentration is out of range
END_VAR

// 段1｜出口预置
FC_DL_ReStripAcidDosageCalc := FALSE;   // 返回值预置假 EN: preset the return value to false
rReMolH := DL_RSD_Z;                    // 摩尔流率预置零 [mol/h] EN: preset the molar flow to zero
rAcidKgH := DL_RSD_Z;                   // 纯酸耗量预置零 [kg/h] EN: preset the acid mass flow to zero
rAcidSolM3h := DL_RSD_Z;                // 酸液流量预置零 [m3/h] EN: preset the acid solution flow to zero
rAcidExcessPct := DL_RSD_Z;             // 富余率预置零 [%] EN: preset the surplus to zero
xConcOk := FALSE;                       // 浓度可行标志预置假 EN: preset the concentration flag to false
xValid := FALSE;                        // 有效标志预置假 EN: preset the validity flag to false
nFaultCode := 0;                        // 故障码预置零 EN: preset the fault code to zero

// 段2｜非有限闸：六个浮点入参全列
xFinAll := (rOrgReConcGpl = rOrgReConcGpl) AND ((rOrgReConcGpl - rOrgReConcGpl) = DL_RSD_Z)
        AND (rFlowOrgM3h = rFlowOrgM3h) AND ((rFlowOrgM3h - rFlowOrgM3h) = DL_RSD_Z)
        AND (rReMolWeight = rReMolWeight) AND ((rReMolWeight - rReMolWeight) = DL_RSD_Z)
        AND (rAcidEquiv = rAcidEquiv) AND ((rAcidEquiv - rAcidEquiv) = DL_RSD_Z)
        AND (rAcidMolWeight = rAcidMolWeight) AND ((rAcidMolWeight - rAcidMolWeight) = DL_RSD_Z)
        AND (rAcidConcGpl = rAcidConcGpl) AND ((rAcidConcGpl - rAcidConcGpl) = DL_RSD_Z);   // 六输入有限性 EN: the finiteness of all six inputs
IF NOT xFinAll THEN                                                                          // 非有限出口 EN: leave early on a non finite input
    nFaultCode := DL_RSD_C_BAD;                                                              // 输入非法码 EN: the illegal input code
    RETURN;                                                                                  // 早退 EN: return early
END_IF

// 段3｜域闸：四个除数逐一过下限（摩尔质量两枚、当量、配酸浓度），流量与浓度非负
IF (rReMolWeight < DL_RSD_MIN) OR (rAcidMolWeight < DL_RSD_MIN)
   OR (rAcidEquiv < DL_RSD_MIN) OR (ABS(rAcidConcGpl) < DL_RSD_MIN)
   OR (rFlowOrgM3h < DL_RSD_Z) OR (rOrgReConcGpl < DL_RSD_Z) THEN
    nFaultCode := DL_RSD_C_RANGE;                                                            // 越域码 EN: the out of range code
    RETURN;                                                                                  // 早退 EN: return early
END_IF

// 段4｜主体：mol/h → 纯酸 kg/h → 酸液 m3/h
rMolH := (rOrgReConcGpl * rFlowOrgM3h * DL_RSD_K1000) / rReMolWeight;                       // 稀土摩尔流率 [mol/h] EN: the rare earth molar flow
rAcidKg := (rMolH * rAcidEquiv * rAcidMolWeight) / DL_RSD_K1000;                             // 纯酸耗量 [kg/h] EN: the pure acid mass flow
rSolM3h := rAcidKg / rAcidConcGpl;                                                           // 酸液体积流量 [m3/h] EN: the acid solution flow, g/L equals kg/m3

// 段5｜结果复检：三路输出非有限或为负一律出口
IF (rMolH <> rMolH) OR (rAcidKg <> rAcidKg) OR (rSolM3h <> rSolM3h)
   OR (rMolH < DL_RSD_Z) OR (rAcidKg < DL_RSD_Z) OR (rSolM3h < DL_RSD_Z) THEN
    nFaultCode := DL_RSD_C_RANGE;                                                            // 复检失败码 EN: the recheck failure code
    RETURN;                                                                                  // 早退，出口保持零哨兵 EN: return early with the zero sentinels
END_IF

// 段6｜浓度校核：同等有机相体积下的供酸能力，不足仅信息级告警
rSupply := rAcidConcGpl * rFlowOrgM3h;                                                       // 同体积供酸能力 [kg/h] EN: the acid supply capability at the same volume
IF (rSupply > DL_RSD_Z) AND (rAcidKg > DL_RSD_MIN) THEN                                       // 供酸能力与酸耗双分母有效 EN: both divisors are usable
    rAcidExcessPct := ((rSupply - rAcidKg) / rAcidKg) * DL_RSD_HUND;                         // 富余率 [%] EN: the surplus percent
    xConcOk := rSupply >= rAcidKg;                                                           // 浓度足以供酸 EN: the concentration is sufficient
ELSE
    rAcidExcessPct := DL_RSD_Z;                                                              // 供酸能力或酸耗为零时给零 [%] EN: give zero when either divisor is zero
    xConcOk := FALSE;                                                                        // 不可供酸 EN: cannot supply
END_IF
rReMolH := rMolH;                                                                            // 摩尔流率出口 [mol/h] EN: the molar flow output
rAcidKgH := rAcidKg;                                                                         // 纯酸耗量出口 [kg/h] EN: the acid mass flow output
rAcidSolM3h := rSolM3h;                                                                      // 酸液流量出口 [m3/h] EN: the acid solution flow output
xValid := TRUE;                                                                              // 结果可信 EN: the results are valid
FC_DL_ReStripAcidDosageCalc := TRUE;                                                         // 返回真 EN: return true
END_FUNCTION

(* ---- FC_DL_ReTheoreticalStagesCalc.st ---- *)
(*
  Component : FC_DL_ReTheoreticalStagesCalc
  Category  : DL_Process
  Function  : 逆流萃取理论级数 n = LN((x0-xStar)/(xn-xStar)) / LN(E)，E 为单级萃取比
  Complexity: C2
  开源溯源 : DLF 内部原创（R94 族模板派生）；参考语义来源见 SOURCE_HUNTING_MATRIX.md
  规则遵从 : R1-R16
  契约     : 输入 rFeedX0 料液浓度 [g/L]、rRaffXn 目标萃余液浓度 [g/L]、rEquilXStar 平衡浓度 [g/L]、
             rExtractRatio 单级萃取比 E [-][>1]；输出 rStages 理论级数 [-]、nStagesCeil 向上取整级数 [级]、
             xValid 有效标志、nFaultCode 故障码；返回 TRUE 表示两输出可信。
  边界     : 须 x0 > xn > xStar；E 须 >1（E≤1 时 LN(E)≤0，理论级数无解，判 9803 并输出无效标志）；
             (x0-xStar) 与 (xn-xStar) 须 >1.0E-9；级数上限 1000，超限判 9804 防 INT 溢出；
             零点五级以下按「先 TRUNC 后按余量进位」向上取整，禁 TRUNC(x)+1。
  码位     : 9801 输入非有限；9802 浓度关系非法；9803 萃取比不足（E≤1）；9804 级数超上限。全部故障级。
*)
FUNCTION FC_DL_ReTheoreticalStagesCalc : BOOL
VAR_INPUT
    rFeedX0       : LREAL := 10.0;   // 料液稀土浓度 x0 [g/L] EN: the rare earth concentration of the feed liquor
    rRaffXn       : LREAL := 0.1;    // 目标萃余液浓度 xn [g/L] EN: the target rare earth concentration of the raffinate
    rEquilXStar   : LREAL := 0.0;    // 平衡浓度 xStar [g/L] EN: the equilibrium concentration of the aqueous phase
    rExtractRatio : LREAL := 3.0;    // 单级萃取比 E，每级浓度下降倍数 [-] EN: the per stage extraction ratio above one
END_VAR
VAR_OUTPUT
    rStages     : LREAL;             // 理论级数（未取整） [级] EN: the theoretical stage number before rounding
    nStagesCeil : INT;               // 向上取整后的工程级数 [级] EN: the engineering stage number rounded upward
    xValid      : BOOL;              // 输出可信标志 EN: the outputs are valid
    nFaultCode  : INT;               // 0=无故障 9801=非有限 9802=浓度关系非法 9803=萃取比不足 9804=级数超限 EN: zero none, 9801 non finite, 9802 illegal concentration order, 9803 ratio too low, 9804 stage overflow
END_VAR
VAR
    xFinAll  : BOOL;                 // 四输入同时有限 EN: all four inputs are finite
    rTopNum  : LREAL;                // 浓度比分子 x0 - x* [g/L] EN: the numerator concentration difference
    rBotNum  : LREAL;                // 浓度比分母 xn - x* [g/L] EN: the denominator concentration difference
    rConcRat : LREAL;                // 浓度比 (x0-xStar)/(xn-xStar) [-] EN: the concentration ratio
    rLnE     : LREAL;                // LN(E) [-] EN: the natural logarithm of the extraction ratio
    rLnRat   : LREAL;                // LN(浓度比) [-] EN: the natural logarithm of the concentration ratio
    rN       : LREAL;                // 理论级数中间值 [级] EN: the interim theoretical stage number
    rTrunc   : LREAL;                // TRUNC 后的整数部分 [级] EN: the truncated integer part
    nCeil    : INT;                  // 进位后的整数级数 [级] EN: the ceiling stage count as an integer
END_VAR
VAR CONSTANT
    DL_RTS_Z       : LREAL := 0.0;    // 浮点零常量 EN: the floating point zero constant
    DL_RTS_ONE     : LREAL := 1.0;    // 浮点壹常量 EN: the floating point one constant
    DL_RTS_EPS     : LREAL := 1.0E-9; // 浓度差与对数的下限 EN: the lower bound of the concentration difference and logarithm
    DL_RTS_STG_MAX : LREAL := 1000.0; // 级数上限（防 INT 溢出） [级] EN: the stage upper bound preventing an integer overflow
    DL_RTS_C_BAD   : INT := 9801;     // 输入非有限 EN: a non finite input
    DL_RTS_C_ORDER : INT := 9802;     // 浓度关系非法 EN: an illegal concentration order
    DL_RTS_C_RATIO : INT := 9803;     // 萃取比不足 EN: the extraction ratio is not above one
    DL_RTS_C_OVER  : INT := 9804;     // 级数超上限 EN: the stage count overflow
END_VAR

// 段1｜出口预置
FC_DL_ReTheoreticalStagesCalc := FALSE;  // 返回值预置假 EN: preset the return value to false
rStages := DL_RTS_Z;                     // 理论级数预置零 [级] EN: preset the theoretical stages to zero
nStagesCeil := 0;                        // 整数级数预置零 [级] EN: preset the integer stages to zero
xValid := FALSE;                         // 有效标志预置假 EN: preset the validity flag to false
nFaultCode := 0;                         // 故障码预置零 EN: preset the fault code to zero

// 段2｜非有限闸：四个浮点入参全部列入，缺一个即对应判据静默失效
xFinAll := (rFeedX0 = rFeedX0) AND ((rFeedX0 - rFeedX0) = DL_RTS_Z)
        AND (rRaffXn = rRaffXn) AND ((rRaffXn - rRaffXn) = DL_RTS_Z)
        AND (rEquilXStar = rEquilXStar) AND ((rEquilXStar - rEquilXStar) = DL_RTS_Z)
        AND (rExtractRatio = rExtractRatio) AND ((rExtractRatio - rExtractRatio) = DL_RTS_Z);   // 四输入有限性 EN: the finiteness of all four inputs
IF NOT xFinAll THEN                                                                              // 非有限出口 EN: leave early on a non finite input
    nFaultCode := DL_RTS_C_BAD;                                                                  // 非有限码 EN: the non finite code
    RETURN;                                                                                      // 早退 EN: return early
END_IF

// 段3｜域闸：浓度关系必须 x0 > xn > x*，否则对数式无物理意义
rTopNum := rFeedX0 - rEquilXStar;                                                               // 分子浓度差 [g/L] EN: the numerator concentration difference
rBotNum := rRaffXn - rEquilXStar;                                                               // 分母浓度差 [g/L] EN: the denominator concentration difference
IF (rTopNum <= DL_RTS_EPS) OR (rBotNum <= DL_RTS_EPS) OR (rTopNum <= rBotNum) THEN              // 浓度顺序与量级闸 EN: the concentration order and magnitude gate
    nFaultCode := DL_RTS_C_ORDER;                                                               // 浓度关系非法码 EN: the illegal concentration order code
    RETURN;                                                                                     // 早退 EN: return early
END_IF

// 段4｜萃取比闸：E 须 >1+容差，E≤1 时理论级数无解（本题明确要求输出无效标志）
IF rExtractRatio <= (DL_RTS_ONE + DL_RTS_EPS) THEN                                              // 萃取比不足闸 EN: the extraction ratio is not above one
    nFaultCode := DL_RTS_C_RATIO;                                                               // 萃取比不足码 EN: the ratio too low code
    RETURN;                                                                                     // 早退 EN: return early
END_IF

// 段5｜主体：n = LN((x0-xStar)/(xn-xStar)) / LN(E)
rConcRat := rTopNum / rBotNum;                                                                  // 浓度比，分母已证 >1.0E-9 [-] EN: the concentration ratio, the denominator is proven positive
rLnRat := LN(rConcRat);                                                                         // 浓度比对数 [-] EN: the logarithm of the concentration ratio
rLnE := LN(rExtractRatio);                                                                      // 萃取比对数，已证 >0 [-] EN: the logarithm of the extraction ratio, proven positive
IF ABS(rLnE) < DL_RTS_EPS THEN                                                                  // 除数下限保护 EN: guard the divisor magnitude
    nFaultCode := DL_RTS_C_RATIO;                                                               // 退化为萃取比不足码 EN: fall back to the ratio code
    RETURN;                                                                                     // 早退 EN: return early
END_IF
rN := rLnRat / rLnE;                                                                            // 理论级数 [级] EN: the theoretical stage number
IF (rN <> rN) OR (rN < DL_RTS_Z) OR (rN > DL_RTS_STG_MAX) THEN                                   // 结果复检：非有限/负/超上限 EN: recheck for a non finite, negative or oversized result
    nFaultCode := DL_RTS_C_OVER;                                                                // 级数超限码 EN: the stage overflow code
    RETURN;                                                                                     // 早退 EN: return early
END_IF

// 段6｜向上取整：先 TRUNC 再按余量进位，整除点不自增（禁 TRUNC(x)+1）
rTrunc := TRUNC(rN);                                                                            // 取整数部分 [级] EN: take the integer part
nCeil := LREAL_TO_INT(rTrunc);                                                                  // 转 INT [级] EN: convert the integer part to an integer
IF rN > rTrunc THEN                                                                             // 余量判据：非整点才进位 EN: only carry when there is a remainder
    IF nCeil < 1000 THEN                                                                        // 进位前上限兜底 EN: bound the carry before it happens
        nCeil := nCeil + 1;                                                                     // 进一级 [级] EN: carry one stage
    END_IF
END_IF
rStages := rN;                                                                                  // 理论级数出口 [级] EN: publish the theoretical stages
nStagesCeil := nCeil;                                                                           // 工程级数出口 [级] EN: publish the engineering stage count
xValid := TRUE;                                                                                 // 结果可信 EN: the results are valid
FC_DL_ReTheoreticalStagesCalc := TRUE;                                                          // 返回真 EN: return true
END_FUNCTION

(* ---- FC_DL_ReWashRatioCalc.st ---- *)
(*
  Component : FC_DL_ReWashRatioCalc
  Category  : DL_Process
  Function  : 洗涤液配比与洗涤级数反算：按杂质夹带率 n = LN(cOut/cIn) / LN(1/(1+R))
  Complexity: C2
  开源溯源 : DLF 内部原创（R94 族模板派生）；参考语义来源见 SOURCE_HUNTING_MATRIX.md
  规则遵从 : R1-R16
  契约     : 输入 rImpInPpm 洗涤前杂质夹带 [ppm]、rImpOutPpm 洗涤后目标杂质 [ppm]、
             rWashRatio 洗涤液与有机相体积配比 W/O [-]、rFlowOrgM3h 有机相流量 [m3/h]；
             输出 rWashFlowM3h 洗涤液体积流量 [m3/h]、rStages 理论洗涤级数 [级]、nStagesCeil 向上取整级数 [级]、
             xValid 有效标志、nFaultCode 故障码。
  边界     : 单级杂质残留比 = 1/(1+R)，故 n = LN(入口/出口) / LN(1+R)；R 须 >1.0E-9、
             入口/出口浓度须 >0 且入口 > 出口，否则判 9802；级数上限 1000 判 9804；
             向上取整先 TRUNC 再按余量进位，整除点不自增。
  码位     : 9801 输入非法（故障级）；9802 浓度或配比关系非法（故障级）；9804 级数超上限（故障级）。
*)
FUNCTION FC_DL_ReWashRatioCalc : BOOL
VAR_INPUT
    rImpInPpm  : LREAL := 500.0;    // 洗涤前杂质夹带量 [ppm] EN: the entrained impurity before washing
    rImpOutPpm : LREAL := 20.0;     // 洗涤后目标杂质含量 [ppm] EN: the target impurity after washing
    rWashRatio : LREAL := 0.3;      // 洗涤液与有机相体积配比 W/O [-] EN: the wash liquid to organic volumetric ratio
    rFlowOrgM3h: LREAL := 5.0;      // 有机相体积流量 [m3/h] EN: the volumetric flow of the organic phase
END_VAR
VAR_OUTPUT
    rWashFlowM3h : LREAL;           // 洗涤液体积流量 [m3/h] EN: the wash liquid volumetric flow
    rStages      : LREAL;           // 理论洗涤级数（未取整） [级] EN: the theoretical wash stage number before rounding
    nStagesCeil  : INT;             // 向上取整后的洗涤级数 [级] EN: the wash stage number rounded upward
    xValid       : BOOL;            // 输出可信标志 EN: the outputs are valid
    nFaultCode   : INT;             // 0=无故障 9801=输入非法 9802=浓度或配比关系非法 9804=级数超上限 EN: zero none, 9801 illegal input, 9802 illegal concentration or ratio, 9804 stage overflow
END_VAR
VAR
    xFinAll  : BOOL;                // 四输入同时有限 EN: all four inputs are finite
    rRatC    : LREAL;               // 进出口杂质浓度比 [-] EN: the inlet to outlet impurity ratio
    rLnC     : LREAL;               // 浓度比对数 [-] EN: the logarithm of the concentration ratio
    rLnR     : LREAL;               // 单级残留系数对数 [-] EN: the logarithm of the single stage retention factor
    rN       : LREAL;               // 级数中间值 [级] EN: the interim stage number
    rTrunc   : LREAL;               // 取整部分 [级] EN: the truncated integer part
    nCeil    : INT;                 // 进位后级数 [级] EN: the ceiling stage count
END_VAR
VAR CONSTANT
    DL_RWR_Z       : LREAL := 0.0;    // 浮点零常量 EN: the floating point zero constant
    DL_RWR_ONE     : LREAL := 1.0;    // 浮点壹常量 EN: the floating point one constant
    DL_RWR_MIN     : LREAL := 1.0E-9; // 浓度与配比的下限 EN: the lower bound of the concentration and the ratio
    DL_RWR_STG_MAX : LREAL := 1000.0; // 级数上限 [级] EN: the stage upper bound
    DL_RWR_C_BAD   : INT := 9801;     // 输入非法 EN: an illegal input
    DL_RWR_C_ORDER : INT := 9802;     // 浓度或配比关系非法 EN: an illegal concentration or ratio order
    DL_RWR_C_OVER  : INT := 9804;     // 级数超上限 EN: the stage count overflow
END_VAR

// 段1｜出口预置
FC_DL_ReWashRatioCalc := FALSE;   // 返回值预置假 EN: preset the return value to false
rWashFlowM3h := DL_RWR_Z;         // 洗涤液流量预置零 [m3/h] EN: preset the wash flow to zero
rStages := DL_RWR_Z;              // 理论级数预置零 [级] EN: preset the theoretical stages to zero
nStagesCeil := 0;                 // 整数级数预置零 [级] EN: preset the integer stages to zero
xValid := FALSE;                  // 有效标志预置假 EN: preset the validity flag to false
nFaultCode := 0;                  // 故障码预置零 EN: preset the fault code to zero

// 段2｜非有限闸：四输入全列
xFinAll := (rImpInPpm = rImpInPpm) AND ((rImpInPpm - rImpInPpm) = DL_RWR_Z)
        AND (rImpOutPpm = rImpOutPpm) AND ((rImpOutPpm - rImpOutPpm) = DL_RWR_Z)
        AND (rWashRatio = rWashRatio) AND ((rWashRatio - rWashRatio) = DL_RWR_Z)
        AND (rFlowOrgM3h = rFlowOrgM3h) AND ((rFlowOrgM3h - rFlowOrgM3h) = DL_RWR_Z);   // 四输入有限性 EN: the finiteness of all four inputs
IF NOT xFinAll THEN                                                                      // 非有限出口 EN: leave early on a non finite input
    nFaultCode := DL_RWR_C_BAD;                                                          // 输入非法码 EN: the illegal input code
    RETURN;                                                                              // 早退 EN: return early
END_IF

// 段3｜域闸：配比与流量为正、出口杂质为正且小于入口，否则对数式无解
IF (rWashRatio < DL_RWR_MIN) OR (rFlowOrgM3h < DL_RWR_Z)
   OR (rImpOutPpm < DL_RWR_MIN) OR (rImpInPpm <= rImpOutPpm) THEN
    nFaultCode := DL_RWR_C_ORDER;                                                        // 关系非法码 EN: the illegal relation code
    RETURN;                                                                              // 早退 EN: return early
END_IF

// 段4｜主体：级数 n = LN(入口/出口) / LN(1+R)
rRatC := rImpInPpm / rImpOutPpm;                                                         // 浓度比，分母已证 >1.0E-9 [-] EN: the concentration ratio, the divisor is proven positive
rLnC := LN(rRatC);                                                                       // 浓度比对数 [-] EN: the logarithm of the concentration ratio
rLnR := LN(DL_RWR_ONE + rWashRatio);                                                     // 单级残留系数对数，已证 >0 [-] EN: the logarithm of the retention factor, proven positive
IF ABS(rLnR) < DL_RWR_MIN THEN                                                           // 除数下限保护 EN: guard the divisor magnitude
    nFaultCode := DL_RWR_C_ORDER;                                                        // 退化为关系非法码 EN: fall back to the relation code
    RETURN;                                                                              // 早退 EN: return early
END_IF
rN := rLnC / rLnR;                                                                       // 洗涤级数 [级] EN: the wash stage number
IF (rN <> rN) OR (rN < DL_RWR_Z) OR (rN > DL_RWR_STG_MAX) THEN                           // 结果复检 EN: recheck the result
    nFaultCode := DL_RWR_C_OVER;                                                         // 级数超限码 EN: the stage overflow code
    RETURN;                                                                              // 早退 EN: return early
END_IF

// 段5｜向上取整：先 TRUNC 再按余量进位
rTrunc := TRUNC(rN);                                                                     // 取整部分 [级] EN: the truncated part
nCeil := LREAL_TO_INT(rTrunc);                                                           // 转 INT [级] EN: convert to an integer
IF rN > rTrunc THEN                                                                      // 余量判据 EN: the remainder test
    IF nCeil < 1000 THEN                                                                 // 进位上限兜底 EN: bound the carry
        nCeil := nCeil + 1;                                                              // 进一级 EN: carry one stage
    END_IF
END_IF
rWashFlowM3h := rWashRatio * rFlowOrgM3h;                                                // 洗涤液流量 [m3/h] EN: the wash liquid flow
rStages := rN;                                                                           // 理论级数出口 [级] EN: the theoretical stages output
nStagesCeil := nCeil;                                                                    // 整数级数出口 [级] EN: the integer stages output
xValid := TRUE;                                                                          // 结果可信 EN: the results are valid
FC_DL_ReWashRatioCalc := TRUE;                                                           // 返回真 EN: return true
END_FUNCTION

(* ---- FC_DL_RinseDragOutCalc.st ---- *)
(*
  DL Factory R83 | FC_DL_RinseDragOutCalc
  功能：由带出液量与浓度差算稀释补水率，并给每小时换槽次数与稳态浓度。
  开源溯源：无（clean-room 自研，依据公开工艺公式，来源=行业通用公式，许可证=MIT，借鉴点=公式结构）
  规则：R1-R21 全遵守
*)
FUNCTION FC_DL_RinseDragOutCalc : REAL
VAR_INPUT
    fDragLph       : REAL; // 工件带出液量 [L/h] / Drag-out volume rate [L/h]
    fRinseVolL     : REAL; // 漂洗槽有效容积 [L] / Rinse tank working volume [L]
    fDragConcPct   : REAL; // 带出液主成分浓度 [%] / Drag-out main component concentration [%]
    fTargetConcPct : REAL; // 漂洗槽允许稳态浓度 [%] / Allowed steady concentration [%]
END_VAR
VAR_OUTPUT
    fDilutionLph : REAL; // 稀释补水率（负值按零）[L/h] / Dilution make-up rate [L/h]
    fTurnsPh     : REAL; // 每小时换槽次数（槽容周转率）[次/h] / Tank turnovers per hour [1/h]
    fSteadyPct   : REAL; // 无补水时稳态平衡浓度 [%] / Steady concentration without make-up [%]
    xValid       : BOOL; // 计算有效性标志 / Calculation validity flag
END_VAR
// 出口预置：四出口统一预置（R256）
fDilutionLph := 0.0; fTurnsPh := 0.0; fSteadyPct := 0.0; xValid := FALSE;
// 非有限拦截 + 量纲自检（R20/R21）
IF NOT (fDragLph > -1.0E30 AND fDragLph < 1.0E30) OR NOT (fRinseVolL > -1.0E30 AND fRinseVolL < 1.0E30) OR NOT (fDragConcPct > -1.0E30 AND fDragConcPct < 1.0E30) OR NOT (fTargetConcPct > -1.0E30 AND fTargetConcPct < 1.0E30) OR fDragLph < 0.0 OR fRinseVolL <= 0.0 OR fDragConcPct <= 0.0 OR fTargetConcPct <= 0.0 THEN
    FC_DL_RinseDragOutCalc := -1.0; RETURN;   // 哨兵 -1：非有限或量纲越界 / Sentinel -1
END_IF
// 浓度次序闸：目标浓度不严于带出浓度时无需稀释
IF fTargetConcPct >= fDragConcPct THEN
    fDilutionLph := 0.0;            // 无需补水 [L/h] / No make-up needed
    fSteadyPct   := fDragConcPct;   // 稳态即带出浓度 [%] / Steady equals drag-out concentration
ELSE
    // 物料平衡：带出带入溶质 = 补水带走溶质，故补水率 = 带出量 × (带出浓度/目标浓度 - 1)
    // 浓度比无量纲，量纲保持 L/h（量纲自洽）
    fDilutionLph := fDragLph * (fDragConcPct / fTargetConcPct - 1.0); // 稀释补水率 [L/h]
    fSteadyPct   := fTargetConcPct; // 补水到位后稳态浓度即目标值 [%] / Steady state hits target
END_IF
// 槽容周转率：L/h ÷ L = 1/h，槽容分母显式零闸（R4/R21）
IF ABS(fRinseVolL) > 1.0E-9 THEN    // 槽容分母显式零闸 / Explicit zero gate on tank volume
    fTurnsPh := fDragLph / fRinseVolL;  // 每小时换槽次数 [次/h] / Tank turnovers per hour
ELSE
    fTurnsPh := 0.0;                // 除零防御缺省 / Divide-by-zero default
END_IF
xValid := TRUE;                             // 链路有效 / Chain valid
FC_DL_RinseDragOutCalc := fDilutionLph;     // 返回稀释补水率 [L/h] / Return dilution rate [L/h]
END_FUNCTION

(* ---- FC_DL_RinseWaterVolumeCalc.st ---- *)
(*
  ============================================================
  组件名 : FC_DL_RinseWaterVolumeCalc
  分类   : DL_Process
  功能   : 冲洗水量计算，由管径管长求管容并按冲洗次数与残留系数折算总耗水量
  复杂度 : C1
  版本   : 1.0.0
  作者   : 道莅工业代码库工厂 / R81
  日期   : 2026-11-24
  开源溯源 : clean-room（no upstream）—— 依据公开工程公式自研，未复制任何上游实现
  红线自检 : R1 无GVL/R2 无物理地址/R3 纯IEC/R4 防除零/R5 双语注释
  接口说明 :
      管容 = pi * (内径/2000)^2 * 管长 * 1000，内径由 mm 先折 m 再折 L，单位链不可省略。
      总水量 = 管容 * 冲洗次数 * (1 + 残留系数)；残留系数限定 0~1。
  ============================================================
*)
FUNCTION FC_DL_RinseWaterVolumeCalc : BOOL
VAR_INPUT
    bEnable       : BOOL; // 使能：TRUE 时计算 / Enable: TRUE to compute
    bErr          : BOOL; // 外部故障：TRUE 时立即退出并置结果无效 / External fault: TRUE aborts with invalid result
    rPipeLen_m    : REAL; // 管道长度 [m] / pipe length [metre]
    rPipeDia_mm   : REAL; // 管道内径 [mm] / pipe inner diameter [millimetre]
    iRinseCount   : INT;  // 冲洗次数 [次] / number of rinse cycles [time]
    rResidFactor  : REAL; // 残留附加系数 [无量纲] / residual surcharge factor [dimensionless]
END_VAR
VAR_OUTPUT
    rPipeVol_L  : REAL; // 单管容积 [L] / single pipe volume [litre]
    rTotalVol_L : REAL; // 全次数冲洗总水量 [L] / total rinse water volume over all cycles [litre]
    bValid      : BOOL; // 输出有效：TRUE 表示结果可用 / Output valid
END_VAR
VAR CONSTANT
    DL_PI      : REAL := 3.14159265; // 圆周率 [无量纲] / circular constant [dimensionless]
    DL_R_MAX   : REAL := 3.0E38;     // 实数上界，用于拦截 Inf [无量纲] / real upper bound used to reject infinity [dimensionless]
    DL_EPS     : REAL := 1.0E-12;    // 除零判定阈值 [无量纲] / division guard threshold [dimensionless]
    DL_MM_TO_M : REAL := 2000.0;     // 直径毫米折半径米的除数 [无量纲] / divisor converting diameter in mm into radius in m [dimensionless]
    DL_M3_TO_L : REAL := 1000.0;     // 立方米折升系数 [L/m3] / cubic metre to litre factor [litre per cubic metre]
    DL_ONE     : REAL := 1.0;        // 单位常量 [无量纲] / unity constant [dimensionless]
    DL_MAX_RINSE : INT := 100;       // 冲洗次数上限 [次] / upper bound of the rinse count [time]
END_VAR
VAR
    _bFin  : BOOL := FALSE; // 输入有限性判定结果 / input finiteness verdict
    _rRad  : REAL := 0.0;   // 管道内半径 [m] / pipe inner radius [metre]
    _rArea : REAL := 0.0;   // 管道过流截面积 [m2] / pipe flow cross section area [square metre]
    _rCnt  : REAL := 0.0;   // 冲洗次数折算实数 [次] / rinse count cast to real [time]
END_VAR

    // 段 1｜出口预置
    rPipeVol_L := 0.0;
    rTotalVol_L := 0.0;
    bValid := FALSE;
    // 段 2｜使能闸与外部故障闸
    IF NOT bEnable THEN
        RETURN;
    END_IF;
    IF bErr THEN
        RETURN;
    END_IF;
    // 段 3｜非有限闸
    _bFin := (rPipeLen_m = rPipeLen_m) AND (ABS(rPipeLen_m) <= DL_R_MAX) AND (rPipeDia_mm = rPipeDia_mm) AND (ABS(rPipeDia_mm) <= DL_R_MAX) AND (rResidFactor = rResidFactor) AND (ABS(rResidFactor) <= DL_R_MAX);
    IF NOT _bFin THEN
        RETURN;
    END_IF;
    // 段 4｜域闸：管长非负、管径严格为正、冲洗次数 1~100、残留系数 0~1
    IF (rPipeLen_m < 0.0) OR (ABS(rPipeDia_mm) <= DL_EPS) OR (rPipeDia_mm < 0.0) THEN
        RETURN;
    END_IF;
    IF (iRinseCount < 1) OR (iRinseCount > DL_MAX_RINSE) THEN
        RETURN;
    END_IF;
    IF (rResidFactor < 0.0) OR (rResidFactor > DL_ONE) THEN
        RETURN;
    END_IF;
    // 段 5｜截面积与单管容积
    _rRad := rPipeDia_mm / DL_MM_TO_M;
    _rArea := DL_PI * _rRad * _rRad;
    rPipeVol_L := _rArea * rPipeLen_m * DL_M3_TO_L;
    // 段 6｜总水量
    _rCnt := INT_TO_REAL(iRinseCount);
    rTotalVol_L := rPipeVol_L * _rCnt * (DL_ONE + rResidFactor);
    bValid := TRUE;
    FC_DL_RinseWaterVolumeCalc := bValid;
END_FUNCTION

(* ---- FC_DL_RoBrineFlowTargetCalc.st ---- *)
(*
  Name: FC_DL_RoBrineFlowTargetCalc
  Category: DL_Process
  Version: 1.0.0
  Round: R90 / 2026-11-25
  开源溯源：clean-room 自研（族 RO/NF 膜法水处理，ST 开源生态实测 0 命中，无外部代码引入）
  功能：1) 按目标回收率反算浓水排放流量的前馈目标值：容积守恒下浓水 = 进水 × (1 − 回收率/100)。
           回收率是「产水占进水的百分比」，故 (1 − 回收率/100) 是「浓水占进水的比例」，
           两者互补且归一化到 0~1，方向固定不可交换（写反会把浓水目标算成产水目标）。
        2) 对反算结果做最小浓水流量下限保护：RO 膜必须维持最低浓水排放以带走盐分并维持横流，
           若反算值低于 fMinBrineFlowM3h，则输出被抬到该下限。此保护是设计动作而非故障，
           故不置 xValid=FALSE；下游若需判别是否被接管，可用
           fFeedFlowM3h × (1 − fTargetRecoveryPct/100) 回算后与 fBrineTargetM3h 比对。
  边界条件：1) 非有限值闸：三路实值入参统一过 NOT(x > -DL_BIG AND x < DL_BIG)，
           同时拦 NaN 与 Inf，命中即拦断实值通路（fBrineTargetM3h 强制 0.0）并置无效（R19）。
        2) 进水流量零闸：ABS(fFeedFlowM3h) > DL_EPS 才允许相乘得到有意义的目标值，
           否则判无效；进水量为负同样判无效（不取 ABS 掩盖反向）。
        3) 目标回收率窄闸：须落在 0.0 ~ 99.99 % 的闭开区间内。回收率 = 100 % 时浓水目标为 0，
           与膜必须维持最小浓水流量的物理事实矛盾，故一律判无效而不输出 0。
        4) 最小浓水流量为负判无效（组态错误）；为 0 表示不设下限保护，属合法组态。
        5) 输出饱和钳制：fBrineTargetM3h 钳到 0 ~ DL_BIG，防极端进水流量导致溢出。
        6) 无回差环节：纯函数无状态，不做迟滞。
  量纲自证：fBrineTargetM3h = (m3/h) × (1 − %/100) = (m3/h) × [-] = m3/h；
           「回收率/100」是无因次归一比例，「1 − 比例」仍为无因次，量纲关系合法。
*)

FUNCTION FC_DL_RoBrineFlowTargetCalc : BOOL
VAR_INPUT
    fFeedFlowM3h        : REAL;   // 系统进水体积流量 [m3/h] / Feed volumetric flow [m3/h]
    fTargetRecoveryPct  : REAL;   // 目标回收率 [%] / Target recovery ratio [%]
    fMinBrineFlowM3h    : REAL;   // 最小浓水排放流量下限 [m3/h] / Minimum brine flow limit [m3/h]
END_VAR
VAR_OUTPUT
    fBrineTargetM3h     : REAL;   // 浓水排放流量目标值 [m3/h] / Brine flow target [m3/h]
    xValid              : BOOL;   // 计算有效标志 [bool] / Calculation valid flag [bool]
END_VAR
VAR
    _fBrineRatio        : REAL;   // 浓水占进水的归一比例 [-] / Brine fraction of feed [-]
    _fBrineRawM3h       : REAL;   // 下限保护前的浓水目标 [m3/h] / Brine target before floor [m3/h]
    _fBrineFloorM3h     : REAL;   // 下限保护后的浓水目标 [m3/h] / Brine target after floor [m3/h]
END_VAR
VAR CONSTANT
    DL_EPS              : REAL := 1.0E-9;   // 分母零闸阈值 [-] / Division-zero gate threshold [-]
    DL_BIG              : REAL := 1.0E12;   // 非有限值闸量级上限 [-] / Finiteness gate magnitude [-]
    DL_PCT              : REAL := 100.0;    // 百分比换算因子 [%] / Percent conversion factor [%]
    DL_REC_OPEN_HI_PCT  : REAL := 99.99;    // 回收率开区间上限 [%] / Recovery open upper bound [%]
END_VAR

(* —— 段 1：非有限值闸（R19：闸断实值通路，NaN 不得乘进目标值） —— *)
IF NOT (fFeedFlowM3h > -DL_BIG AND fFeedFlowM3h < DL_BIG)
   OR NOT (fTargetRecoveryPct > -DL_BIG AND fTargetRecoveryPct < DL_BIG)
   OR NOT (fMinBrineFlowM3h > -DL_BIG AND fMinBrineFlowM3h < DL_BIG) THEN
    fBrineTargetM3h := 0.0;                 // 输出强制 0.0 / Output forced to zero
    xValid := FALSE;                        // 有效位清零 / Validity cleared
    FC_DL_RoBrineFlowTargetCalc := FALSE;   // 返回码同源 / Return mirrors validity
    RETURN;                                 // 立即退出 / Immediate exit
END_IF

(* —— 段 2：进水零闸（R4：容积基准量为 0 则目标值无意义） —— *)
IF ABS(fFeedFlowM3h) <= DL_EPS THEN
    fBrineTargetM3h := 0.0;                 // 输出强制 0.0 / Output forced to zero
    xValid := FALSE;                        // 判无效 / Invalid
    FC_DL_RoBrineFlowTargetCalc := FALSE;   // 返回码同步 / Return synchronised
    RETURN;                                 // 提前退出 / Early exit
END_IF

(* —— 段 3：主算式（R22 方向自核：1 − 回收率/100 是浓水比例，不是产水比例） —— *)
_fBrineRatio := 1.0 - fTargetRecoveryPct / DL_PCT;              // 浓水占比 [-]
_fBrineRawM3h := fFeedFlowM3h * _fBrineRatio;                   // 反算浓水目标 [m3/h]

(* —— 段 4：最小浓水流量下限保护（设计动作，抬高到下限，不判无效） —— *)
_fBrineFloorM3h := MAX(_fBrineRawM3h, fMinBrineFlowM3h);        // 取反算值与下限的较大者 [m3/h]

(* —— 段 5：有效位单点聚合（进水为正 + 回收率窄闸 + 下限组态合法） —— *)
xValid := (fFeedFlowM3h > DL_EPS)                               // 进水必须为正
          AND (fTargetRecoveryPct >= 0.0)                       // 回收率不越下限
          AND (fTargetRecoveryPct <= DL_REC_OPEN_HI_PCT)        // 回收率不得达 100 %
          AND (fMinBrineFlowM3h >= 0.0);                        // 最小浓水流量不得为负

(* —— 段 6：输出单点写盘（饱和钳制后写，禁同拍二次赋值） —— *)
fBrineTargetM3h := LIMIT(0.0, _fBrineFloorM3h, DL_BIG);         // 浓水目标钳 0..DL_BIG [m3/h]
FC_DL_RoBrineFlowTargetCalc := xValid;                          // 返回码：TRUE = 计算可信

END_FUNCTION

(* ---- FC_DL_RoConcentrationPolarizationCalc.st ---- *)
(*
  Name: FC_DL_RoConcentrationPolarizationCalc
  Category: DL_Process
  Version: 1.0.0
  Round: R90 / 2026-11-25
  开源溯源：clean-room 自研（族 RO/NF 膜法水处理，ST 开源生态实测 0 命中，无外部代码引入）
  功能：1) 浓差极化因子按边界层膜模型 β = EXP(J / k) 估算：J 为膜通量换算成的渗透速度（m/s），
           k 为传质系数（m/s），J/k 为无因次的 Péclet 数；β 表示膜面盐浓度相对主体浓度的倍数，
           β 越大结垢与通量衰减风险越高。
        2) 通量入参按工程单位 LMH 接收，先做 LMH → m/s 的两级换算（/1000 L/m3、/3600 s/h），
           保证与传质系数同量纲后才能相除，禁止 LMH 与 m/s 直接相除。
        3) 膜面横流速度参与可行性判定而非进入算式：横流速度是传质系数 k 的物理来源，
           实测横流为零意味着 k 的标定前提失效（层流边界层崩溃），此时 β 模型不可信，
           故对横流做零闸并判无效，而不是把横流再乘一次导致双重计入。
  边界条件：1) 非有限值闸：三路实值入参统一过 NOT(x > -DL_BIG AND x < DL_BIG)，
           同时拦 NaN 与 Inf，命中即拦断实值通路（fCpFactor 强制 0.0）并置无效（R19）。
        2) 传质系数零闸：ABS(fMassTransCoef) > DL_EPS 才允许相除，否则判无效。
        3) 横流速度零闸：fCrossFlowMps <= DL_EPS 判无效（无横流即无稳定边界层）。
        4) Péclet 数上限保护：J/k 先钳到 0 ~ LN(DL_CP_MAX)，防止 EXP 溢出成 Inf；
           β 结果再饱和钳到 DL_CP_MIN ~ DL_CP_MAX（1.0 ~ 3.0），超出即无物理意义。
        5) 通量为负判无效（传感器反向）；通量为 0 属合法工况，β 退化为 1.0。
        6) 无回差环节：纯函数无状态，不做迟滞。
  量纲自证：J = (L/(m2·h)) / 1000 (L/m3) / 3600 (s/h) = m/s；
           J / k = (m/s) / (m/s) = 无因次 Péclet 数 [-]；
           β = EXP([-]) = 无因次浓度比 [-]。
*)

FUNCTION FC_DL_RoConcentrationPolarizationCalc : BOOL
VAR_INPUT
    fFluxLMH         : REAL;   // 膜通量 [L/(m2·h)] / Membrane flux [LMH]
    fCrossFlowMps    : REAL;   // 膜面横流速度 [m/s] / Membrane cross-flow velocity [m/s]
    fMassTransCoef   : REAL;   // 传质系数 k [m/s] / Mass transfer coefficient [m/s]
END_VAR
VAR_OUTPUT
    fCpFactor        : REAL;   // 浓差极化因子 β [-] / Concentration polarization factor [-]
    xValid           : BOOL;   // 计算有效标志 [bool] / Calculation valid flag [bool]
END_VAR
VAR
    _fFluxMps        : REAL;   // 换算后的渗透速度 [m/s] / Permeate velocity [m/s]
    _fPeclet         : REAL;   // Péclet 数 J/k [-] / Peclet number [-]
    _fPecletMax      : REAL;   // Péclet 数上限（由 β 上限反算）[-] / Peclet ceiling [-]
    _fBetaRaw        : REAL;   // 未饱和的极化因子 [-] / Raw polarization factor [-]
END_VAR
VAR CONSTANT
    DL_EPS           : REAL := 1.0E-9;    // 分母零闸阈值 [-] / Division-zero gate threshold [-]
    DL_BIG           : REAL := 1.0E12;    // 非有限值闸量级上限 [-] / Finiteness gate magnitude [-]
    DL_L_PER_M3      : REAL := 1000.0;    // m3 → L 换算因子 [L/m3] / Cubic metre to litre factor [L/m3]
    DL_S_PER_H       : REAL := 3600.0;    // h → s 换算因子 [s/h] / Hour to second factor [s/h]
    DL_CP_MIN        : REAL := 1.0;       // 极化因子饱和下限 [-] / Polarization factor low [-]
    DL_CP_MAX        : REAL := 3.0;       // 极化因子饱和上限 [-] / Polarization factor high [-]
END_VAR

(* —— 段 1：非有限值闸（R19：闸断实值通路，NaN 不进 EXP） —— *)
IF NOT (fFluxLMH > -DL_BIG AND fFluxLMH < DL_BIG)
   OR NOT (fCrossFlowMps > -DL_BIG AND fCrossFlowMps < DL_BIG)
   OR NOT (fMassTransCoef > -DL_BIG AND fMassTransCoef < DL_BIG) THEN
    fCpFactor := 0.0;                       // 输出强制 0.0 / Output forced to zero
    xValid := FALSE;                        // 有效位清零 / Validity cleared
    FC_DL_RoConcentrationPolarizationCalc := FALSE;   // 返回码同源 / Return mirrors validity
    RETURN;                                 // 立即退出 / Immediate exit
END_IF

(* —— 段 2：传质系数零闸 + 横流零闸（R4：两个分母/前提都要闸） —— *)
IF (ABS(fMassTransCoef) <= DL_EPS) OR (fCrossFlowMps <= DL_EPS) THEN
    fCpFactor := 0.0;                       // 前提失效即不给数 / No premise, no number
    xValid := FALSE;                        // 判无效 / Invalid
    FC_DL_RoConcentrationPolarizationCalc := FALSE;   // 返回码同步 / Return synchronised
    RETURN;                                 // 提前退出 / Early exit
END_IF

(* —— 段 3：通量单位换算（LMH → m/s，两级因子不可省略） —— *)
_fFluxMps := MAX(0.0, fFluxLMH) / DL_L_PER_M3 / DL_S_PER_H;   // 渗透速度 [m/s]

(* —— 段 4：Péclet 数与上限保护（先钳指数再 EXP，防溢出成 Inf） —— *)
_fPecletMax := LN(DL_CP_MAX);                                  // 由 β 上限反算的指数上限 [-]
_fPeclet := LIMIT(0.0, _fFluxMps / fMassTransCoef, _fPecletMax);   // J/k 钳 0..LN(3)
_fBetaRaw := EXP(_fPeclet);                                    // 极化因子 [-]

(* —— 段 5：有效位单点聚合（通量非负 + 前提量正） —— *)
xValid := (fFluxLMH >= 0.0)                                    // 通量不得为负
          AND (fMassTransCoef > DL_EPS)                        // 传质系数必须为正
          AND (fCrossFlowMps > DL_EPS);                        // 横流必须为正

(* —— 段 6：输出单点写盘（β 饱和钳到物理域） —— *)
fCpFactor := LIMIT(DL_CP_MIN, _fBetaRaw, DL_CP_MAX);           // β 钳 1.0..3.0 [-]
FC_DL_RoConcentrationPolarizationCalc := xValid;               // 返回码：TRUE = 计算可信

END_FUNCTION

(* ---- FC_DL_RoFluxCalc.st ---- *)
(*
  Name: FC_DL_RoFluxCalc
  Category: DL_Process
  Version: 1.0.0
  Round: R90 / 2026-11-25
  开源溯源：clean-room 自研（族 RO/NF 膜法水处理，ST 开源生态实测 0 命中，无外部代码引入）
  功能：1) 膜通量按「单位时间单位膜面积的产水容积」计算，容积流量由 m3/h 换算为 L/h 后除以面积，
           得 LMH（L/(m2·h)）：fFluxLMH = fPermeateFlowM3h * 1000 / fMembraneAreaM2 * 1，
           其中 1000 为 m3 → L 的换算因子，除的是有效膜面积而非单支膜面积。
        2) 温度校正通量按 25 °C 基准折算：TCF = EXP(LN(DL_TCF_BASE) * (DL_T_REF_C - fTempC))，
           即每偏离基准温度 1 °C 通量按 DL_TCF_BASE 倍率变化；fFluxTempCorrLMH = fFluxLMH * TCF。
           该式用于把不同水温下的通量拉到同一基准比较，禁止直接用实测通量做趋势判定。
  边界条件：1) 面积零闸：ABS(fMembraneAreaM2) > DL_EPS 才允许除法，否则清零输出并置无效。
        2) 非有限值闸：三路实值入参统一过 NOT(x > -DL_BIG AND x < DL_BIG)，同时拦 NaN 与 Inf，
           命中即拦断实值通路（两个 REAL 输出强制 0.0），不许把 NaN 透传（R19）。
        3) 温度量程窄闸：fTempC 须在 DL_T_LO_C..DL_T_HI_C（0 ~ 80 °C）内，越域判无效，
           因为温度校正式的适用域只在膜系统实际水温区间；越域仍按边界值算出一个数供参考。
        4) 通量不得为负：产水流量为负判传感器反向，置无效。
        5) 校正通量做饱和硬限：TCF 结果钳到 0.05 ~ 20.0（对应约 0.5 ~ 25 °C 的极端偏离），
           防止极端温度把校正值放大到无物理意义的量级。
  量纲自证：fFluxLMH = (m3/h) * 1000 (L/m3) / (m2) = L/(m2·h) = LMH，量纲闭合；
           TCF = [-]（无因次倍率），fFluxTempCorrLMH = (L/(m2·h)) * [-] = L/(m2·h)，同量纲。
*)

FUNCTION FC_DL_RoFluxCalc : BOOL
VAR_INPUT
    fPermeateFlowM3h : REAL;   // 产水体积流量 [m3/h] / Permeate volumetric flow [m3/h]
    fMembraneAreaM2  : REAL;   // 有效膜面积 [m2] / Effective membrane area [m2]
    fTempC           : REAL;   // 给水温度 [°C] / Feed water temperature [°C]
END_VAR
VAR_OUTPUT
    fFluxLMH         : REAL;   // 实测膜通量 [L/(m2·h)] / Measured membrane flux [LMH]
    fFluxTempCorrLMH : REAL;   // 25 °C 基准校正通量 [L/(m2·h)] / Temperature-corrected flux [LMH]
    xValid           : BOOL;   // 计算有效标志 [bool] / Calculation valid flag [bool]
END_VAR
VAR
    _fTcf            : REAL;   // 温度校正因子 [-] / Temperature correction factor [-]
    _fTClampedC      : REAL;   // 钳制到适用域内的温度 [°C] / Temperature clamped to valid range [°C]
    _fFluxRawLMH     : REAL;   // 未钳制的原始通量 [L/(m2·h)] / Raw flux before limiting [LMH]
END_VAR
VAR CONSTANT
    DL_EPS           : REAL := 1.0E-9;    // 分母零闸阈值 [-] / Division-zero gate threshold [-]
    DL_BIG           : REAL := 1.0E12;    // 非有限值闸量级上限 [-] / Finiteness gate magnitude [-]
    DL_L_PER_M3      : REAL := 1000.0;    // m3 → L 换算因子 [L/m3] / Cubic metre to litre factor [L/m3]
    DL_T_REF_C       : REAL := 25.0;      // 通量基准温度 [°C] / Flux reference temperature [°C]
    DL_TCF_BASE      : REAL := 1.03;      // 每 °C 通量变化倍率 [-] / Flux change ratio per degC [-]
    DL_T_LO_C        : REAL := 0.0;       // 温度适用域下限 [°C] / Temperature validity low [°C]
    DL_T_HI_C        : REAL := 80.0;      // 温度适用域上限 [°C] / Temperature validity high [°C]
    DL_TCF_MIN       : REAL := 0.05;      // 校正因子饱和下限 [-] / TCF saturation low [-]
    DL_TCF_MAX       : REAL := 20.0;      // 校正因子饱和上限 [-] / TCF saturation high [-]
END_VAR

(* —— 段 1：非有限值闸（R19：同时拦 NaN 与 Inf，并闸断两个 REAL 输出通路） —— *)
IF NOT (fPermeateFlowM3h > -DL_BIG AND fPermeateFlowM3h < DL_BIG)
   OR NOT (fMembraneAreaM2 > -DL_BIG AND fMembraneAreaM2 < DL_BIG)
   OR NOT (fTempC > -DL_BIG AND fTempC < DL_BIG) THEN
    fFluxLMH := 0.0;                        // 输出强制 0.0 / Output forced to zero
    fFluxTempCorrLMH := 0.0;                // 校正通量强制 0.0 / Corrected flux forced to zero
    xValid := FALSE;                        // 有效位清零 / Validity cleared
    FC_DL_RoFluxCalc := FALSE;              // 返回码同源 / Return mirrors validity
    RETURN;                                 // 立即退出 / Immediate exit
END_IF

(* —— 段 2：面积零闸（R4：分母先过 ABS 闸） —— *)
IF ABS(fMembraneAreaM2) <= DL_EPS THEN
    fFluxLMH := 0.0;                        // 无面积即无通量 / No area means no flux
    fFluxTempCorrLMH := 0.0;                // 校正通量同样清零 / Corrected flux cleared
    xValid := FALSE;                        // 判无效 / Invalid
    FC_DL_RoFluxCalc := FALSE;              // 返回码同步 / Return synchronised
    RETURN;                                 // 提前退出 / Early exit
END_IF

(* —— 段 3：实测通量（R22 方向自核：分子为产水容积，分母为膜面积，不取倒数） —— *)
_fFluxRawLMH := fPermeateFlowM3h * DL_L_PER_M3 / fMembraneAreaM2;   // [L/(m2·h)]

(* —— 段 4：温度校正因子（EXPT 的跨平台安全写法：EXP(LN(base) * 指数)） —— *)
_fTClampedC := LIMIT(DL_T_LO_C, fTempC, DL_T_HI_C);                 // 钳到适用域 [°C]
_fTcf := EXP(LN(DL_TCF_BASE) * (DL_T_REF_C - _fTClampedC));         // 25 °C 基准折算 [-]
_fTcf := LIMIT(DL_TCF_MIN, _fTcf, DL_TCF_MAX);                      // 因子饱和硬限 [-]

(* —— 段 5：有效位单点聚合（物理域 + 温度量程 + 非负） —— *)
xValid := (fPermeateFlowM3h >= 0.0)                                 // 产水不得为负
          AND (fMembraneAreaM2 > DL_EPS)                            // 面积必须为正
          AND (fTempC >= DL_T_LO_C)                                 // 温度不越下限
          AND (fTempC <= DL_T_HI_C);                                // 温度不越上限

(* —— 段 6：输出单点写盘（饱和后再写，禁同拍二次赋值） —— *)
fFluxLMH := MAX(0.0, _fFluxRawLMH);                                 // 通量钳 >= 0 [L/(m2·h)]
fFluxTempCorrLMH := MAX(0.0, _fFluxRawLMH * _fTcf);                 // 校正通量钳 >= 0 [L/(m2·h)]
FC_DL_RoFluxCalc := xValid;                                         // 返回码：TRUE = 计算可信

END_FUNCTION

(* ---- FC_DL_RoNetDrivingPressureCalc.st ---- *)
(*
  Name: FC_DL_RoNetDrivingPressureCalc
  Category: DL_Process
  Version: 1.0.0
  Round: R90 / 2026-11-25
  开源溯源：clean-room 自研（族 RO/NF 膜法水处理，ST 开源生态实测 0 命中，无外部代码引入）
  功能：1) 净驱动压按「推动水穿过膜的有效压差」计算，工程口径为
           NDP = (给水压力 + 浓水压力) / 2 − 渗透压 − 浓水侧流道压降。
           平均给水压取首末端两点的算术均值（膜元件内压力沿线近似线性下降），
           减渗透压扣除浓水侧的化学势反压，再减流道压降扣除沿程损失。
        2) NDP <= 0 表示驱动力消失，膜段无法产水（且存在浓差极化与结垢风险），
           判失效并输出 0.0，禁止输出负的驱动压给下游做乘法（会翻转通量符号）。
  边界条件：1) 非有限值闸：四路实值入参统一过 NOT(x > -DL_BIG AND x < DL_BIG)，
           同时拦 NaN 与 Inf，命中即拦断实值通路（fNdpBar 强制 0.0）并置无效（R19）。
        2) 压力量程窄闸 0 ~ DL_P_BAR_MAX（0 ~ 120 bar）：单点越域判无效（变送器故障或超量程），
           越域值钳到量程边界后再参与运算，避免单点异常把 NDP 拉成极端值。
        3) 负压判定：任一路表压为负判无效（RO 系统不允许负压，负压意味着抽真空或量程零点漂移）。
        4) NDP <= 0 判无效并输出 0.0（驱动力消失，非数值问题而是工艺失效）。
        5) 无回差环节：纯函数无状态，迟滞由下游报警件承担。
  量纲自证：fNdpBar = (bar + bar)/2 − bar − bar = bar，四项全部为 bar，量纲一致；
           平均值为 (P_feed + P_conc) / 2，除数 2 是无因次算术平均点数，不引入量纲。
*)

FUNCTION FC_DL_RoNetDrivingPressureCalc : BOOL
VAR_INPUT
    fFeedBar          : REAL;   // 给水侧压力 [bar] / Feed side pressure [bar]
    fConcentrateBar   : REAL;   // 浓水侧压力 [bar] / Concentrate side pressure [bar]
    fOsmoticBar       : REAL;   // 渗透压（已按给水/浓水均值折算）[bar] / Osmotic pressure [bar]
    fChannelDropBar   : REAL;   // 浓水侧流道压降 [bar] / Concentrate channel pressure drop [bar]
END_VAR
VAR_OUTPUT
    fNdpBar           : REAL;   // 净驱动压 [bar] / Net driving pressure [bar]
    xValid            : BOOL;   // 计算有效标志 [bool] / Calculation valid flag [bool]
END_VAR
VAR
    _fFeedClampBar    : REAL;   // 钳制后的给水压力 [bar] / Clamped feed pressure [bar]
    _fConcClampBar    : REAL;   // 钳制后的浓水压力 [bar] / Clamped concentrate pressure [bar]
    _fOsmClampBar     : REAL;   // 钳制后的渗透压 [bar] / Clamped osmotic pressure [bar]
    _fDropClampBar    : REAL;   // 钳制后的流道压降 [bar] / Clamped channel pressure drop [bar]
    _fMeanFeedBar     : REAL;   // 首末端平均给水压力 [bar] / Mean feed pressure [bar]
    _fNdpRawBar       : REAL;   // 未饱和的原始净驱动压 [bar] / Raw NDP before limiting [bar]
END_VAR
VAR CONSTANT
    DL_EPS            : REAL := 1.0E-9;   // 分母零闸阈值 [-] / Division-zero gate threshold [-]
    DL_BIG            : REAL := 1.0E12;   // 非有限值闸量级上限 [-] / Finiteness gate magnitude [-]
    DL_P_BAR_MAX      : REAL := 120.0;    // 压力变送器量程上限 [bar] / Pressure transmitter span high [bar]
    DL_MEAN_POINTS    : REAL := 2.0;      // 平均给水压的取点数 [-] / Averaging point count [-]
END_VAR

(* —— 段 1：非有限值闸（R19：四路入参全覆盖，拦 NaN 与 Inf） —— *)
IF NOT (fFeedBar > -DL_BIG AND fFeedBar < DL_BIG)
   OR NOT (fConcentrateBar > -DL_BIG AND fConcentrateBar < DL_BIG)
   OR NOT (fOsmoticBar > -DL_BIG AND fOsmoticBar < DL_BIG)
   OR NOT (fChannelDropBar > -DL_BIG AND fChannelDropBar < DL_BIG) THEN
    fNdpBar := 0.0;                         // 输出强制 0.0 / Output forced to zero
    xValid := FALSE;                        // 有效位清零 / Validity cleared
    FC_DL_RoNetDrivingPressureCalc := FALSE;   // 返回码同源 / Return mirrors validity
    RETURN;                                 // 立即退出 / Immediate exit
END_IF

(* —— 段 2：负压闸（RO 系统不允许负表压：抽真空或零点漂移均为故障） —— *)
IF (fFeedBar < 0.0) OR (fConcentrateBar < 0.0) OR (fOsmoticBar < 0.0) OR (fChannelDropBar < 0.0) THEN
    fNdpBar := 0.0;                         // 输出强制 0.0 / Output forced to zero
    xValid := FALSE;                        // 判无效 / Invalid
    FC_DL_RoNetDrivingPressureCalc := FALSE;   // 返回码同步 / Return synchronised
    RETURN;                                 // 提前退出 / Early exit
END_IF

(* —— 段 3：量程钳制（单点越量程钳到边界，避免异常点污染整式） —— *)
_fFeedClampBar := LIMIT(0.0, fFeedBar, DL_P_BAR_MAX);            // 给水压力钳 [bar]
_fConcClampBar := LIMIT(0.0, fConcentrateBar, DL_P_BAR_MAX);     // 浓水压力钳 [bar]
_fOsmClampBar := LIMIT(0.0, fOsmoticBar, DL_P_BAR_MAX);          // 渗透压钳 [bar]
_fDropClampBar := LIMIT(0.0, fChannelDropBar, DL_P_BAR_MAX);     // 流道压降钳 [bar]

(* —— 段 4：主算式（R22 方向自核：先平均值，再逐项扣减，扣减项全部为正相加） —— *)
_fMeanFeedBar := (_fFeedClampBar + _fConcClampBar) / DL_MEAN_POINTS;   // 算术均值 [bar]
_fNdpRawBar := _fMeanFeedBar - _fOsmClampBar - _fDropClampBar;         // 净驱动压 [bar]

(* —— 段 5：有效位单点聚合（量程 + 驱动力存在性） —— *)
xValid := (fFeedBar <= DL_P_BAR_MAX)                            // 给水不越量程
          AND (fConcentrateBar <= DL_P_BAR_MAX)                 // 浓水不越量程
          AND (fOsmoticBar <= DL_P_BAR_MAX)                     // 渗透压不越量程
          AND (fChannelDropBar <= DL_P_BAR_MAX)                 // 流道压降不越量程
          AND (_fNdpRawBar > 0.0);                              // 驱动力必须严格为正

(* —— 段 6：输出单点写盘（负值不得流出，否则下游乘法会翻转通量符号） —— *)
fNdpBar := MAX(0.0, _fNdpRawBar);                               // 净驱动压钳 >= 0 [bar]
FC_DL_RoNetDrivingPressureCalc := xValid;                       // 返回码：TRUE = 计算可信

END_FUNCTION

(* ---- FC_DL_RoOsmoticPressureCalc.st ---- *)
(*
  Name: FC_DL_RoOsmoticPressureCalc
  Category: DL_Process
  Version: 1.0.0
  Round: R90 / 2026-11-25
  开源溯源：clean-room 自研（族 RO/NF 膜法水处理，ST 开源生态实测 0 命中，无外部代码引入）
  功能：1) 按 van't Hoff 简化式计算给水渗透压：π = i · C · R · T，其中溶质按 NaCl 双离子
           （i = 2）、摩尔质量折算并入常数项，得到工程式 π[Pa] = DL_VANT_HOFF · T[K] · TDS[mg/L]，
           再除 1.0E5 转 bar；温度以开尔文参与，故必须先做 °C → K 的偏移。
        2) TDS 先做量程钳制（0 ~ DL_TDS_MAX mg/L）再进算式，超域值不让其把渗透压推到无物理意义量级；
           钳制动作本身不置无效，只有负值或非有限才判无效。
  边界条件：1) 非有限值闸：两路实值入参先过 NOT(x > -DL_BIG AND x < DL_BIG)，同时拦 NaN 与 Inf，
           命中即拦断实值通路（fOsmoticBar 强制 0.0）并置 xValid=FALSE（R19）。
        2) TDS 负值判无效（浓度不可能为负，属变送器故障），不取绝对值掩盖。
        3) TDS 上限饱和钳制 DL_TDS_MAX = 60000 mg/L（覆盖海水级高盐工况），超限钳到上限并判无效；
           下限钳 0.0（纯水渗透压为 0，属合法工况，不判无效）。
        4) 温度量程窄闸 0 ~ 90 °C：水温越域钳到边界算参考值并置无效，因为开尔文偏移在负温度附近
           会使简化式显著偏离实测渗透压。
        5) 无回差环节：纯函数无状态，不做迟滞。
  量纲自证：DL_VANT_HOFF = 0.28451 Pa·L/(mg·K)，故 Pa·L/(mg·K) × K × mg/L = Pa，量纲闭合；
           fOsmoticBar = Pa / 1.0E5 (Pa/bar) = bar。
*)

FUNCTION FC_DL_RoOsmoticPressureCalc : BOOL
VAR_INPUT
    fTdsMgL      : REAL;   // 给水总溶解固体 [mg/L] / Feed total dissolved solids [mg/L]
    fTempC       : REAL;   // 给水温度 [°C] / Feed water temperature [°C]
END_VAR
VAR_OUTPUT
    fOsmoticBar  : REAL;   // 给水渗透压 [bar] / Feed osmotic pressure [bar]
    xValid       : BOOL;   // 计算有效标志 [bool] / Calculation valid flag [bool]
END_VAR
VAR
    _fTdsClamp   : REAL;   // 钳制到量程内的 TDS [mg/L] / TDS clamped into range [mg/L]
    _fTClampC    : REAL;   // 钳制到量程内的温度 [°C] / Temperature clamped into range [°C]
    _fTKelvin    : REAL;   // 绝对温度 [K] / Absolute temperature [K]
    _fOsmPa      : REAL;   // 渗透压中间量 [Pa] / Osmotic pressure intermediate [Pa]
END_VAR
VAR CONSTANT
    DL_EPS       : REAL := 1.0E-9;    // 分母零闸阈值 [-] / Division-zero gate threshold [-]
    DL_BIG       : REAL := 1.0E12;    // 非有限值闸量级上限 [-] / Finiteness gate magnitude [-]
    DL_K0        : REAL := 273.15;    // 摄氏转开尔文偏移 [K] / Celsius to Kelvin offset [K]
    DL_VANT_HOFF : REAL := 0.28451;   // van't Hoff 合并常数 [Pa·L/(mg·K)] / Lumped van't Hoff constant
    DL_PA_PER_BAR: REAL := 1.0E5;     // Pa → bar 换算因子 [Pa/bar] / Pascal to bar factor [Pa/bar]
    DL_TDS_MAX   : REAL := 60000.0;   // TDS 量程上限（饱和钳制点）[mg/L] / TDS saturation ceiling [mg/L]
    DL_T_LO_C    : REAL := 0.0;       // 温度量程下限 [°C] / Temperature range low [°C]
    DL_T_HI_C    : REAL := 90.0;      // 温度量程上限 [°C] / Temperature range high [°C]
END_VAR

(* —— 段 1：非有限值闸（R19：闸断实值通路，NaN 不得进入乘加链） —— *)
IF NOT (fTdsMgL > -DL_BIG AND fTdsMgL < DL_BIG)
   OR NOT (fTempC > -DL_BIG AND fTempC < DL_BIG) THEN
    fOsmoticBar := 0.0;                     // 输出强制 0.0 / Output forced to zero
    xValid := FALSE;                        // 有效位清零 / Validity cleared
    FC_DL_RoOsmoticPressureCalc := FALSE;   // 返回码同源 / Return mirrors validity
    RETURN;                                 // 立即退出 / Immediate exit
END_IF

(* —— 段 2：TDS 负值闸（浓度不可为负 = 变送器故障，不取 ABS 掩盖） —— *)
IF fTdsMgL < 0.0 THEN
    fOsmoticBar := 0.0;                     // 输出强制 0.0 / Output forced to zero
    xValid := FALSE;                        // 判无效 / Invalid
    FC_DL_RoOsmoticPressureCalc := FALSE;   // 返回码同步 / Return synchronised
    RETURN;                                 // 提前退出 / Early exit
END_IF

(* —— 段 3：量程钳制（饱和硬限，TDS 上限 / 温度双边界） —— *)
_fTdsClamp := LIMIT(0.0, fTdsMgL, DL_TDS_MAX);        // TDS 钳 0..60000 [mg/L]
_fTClampC := LIMIT(DL_T_LO_C, fTempC, DL_T_HI_C);     // 温度钳 0..90 [°C]
_fTKelvin := _fTClampC + DL_K0;                       // °C → K [K]

(* —— 段 4：van't Hoff 简化式（R22 方向自核：乘温度、乘浓度，均为正相关） —— *)
_fOsmPa := DL_VANT_HOFF * _fTKelvin * _fTdsClamp;     // 渗透压 [Pa]

(* —— 段 5：有效位单点聚合（越量程判无效，钳制值仍输出供参考） —— *)
xValid := (fTdsMgL <= DL_TDS_MAX)                     // TDS 不越上限
          AND (fTempC >= DL_T_LO_C)                   // 温度不越下限
          AND (fTempC <= DL_T_HI_C);                  // 温度不越上限

(* —— 段 6：输出单点写盘（Pa → bar，饱和保护防溢出） —— *)
fOsmoticBar := LIMIT(0.0, _fOsmPa / DL_PA_PER_BAR, DL_BIG);   // 渗透压钳 0..DL_BIG [bar]
FC_DL_RoOsmoticPressureCalc := xValid;                        // 返回码：TRUE = 计算可信

END_FUNCTION
